// TIA Portal project "环氧乙烷灭菌器（XG2-C）260909_V18" (V18)

(* hardware
DEVICE "S7-1200 station_1"  S7-1200 Station
   slot 0: "Rack_0"  S7-1200 Rack  Rack  V1.0
   slot 1: "PLC_1"  CPU 1214C DC/DC/DC  6ES7 214-1AG40-0XB0  V4.2
   slot 2: "DI 8x24VDC_1"  6ES7 221-1BF32-0XB0  V2.0
   slot 3: "DQ 8x24VDC _1"  SM 1222 DQ8 x 24VDC  6ES7 222-1BF32-0XB0  V2.0
   slot 4: "DQ 8x24VDC _2"  SM 1222 DQ8 x 24VDC  6ES7 222-1BF32-0XB0  V2.0
   slot 5: "AI 4xRTD_1"  SM 1231 AI4 x RTD  6ES7 231-5PD32-0XB0  V2.0
   slot 6: "AI 4x13BIT_1"  6ES7 231-4HD32-0XB0  V2.0
*)

// ===== PLC "PLC_1"  CPU 1214C DC/DC/DC =====
// protected blocks, not shown: "0程序运行控制流程", "1预处理", "2保压", "3加湿", "4加药", "5灭菌", "6脉动", "7通风", "Main", "紧急脉动", "紧急通风"

VAR_GLOBAL   // PLC tag table "默认变量表"
   "Clock_Byte" AT %MB0 : Byte;
   "Clock_10Hz" AT %M0.0 : Bool;
   "Clock_5Hz" AT %M0.1 : Bool;
   "Clock_2.5Hz" AT %M0.2 : Bool;
   "Clock_2Hz" AT %M0.3 : Bool;
   "Clock_1.25Hz" AT %M0.4 : Bool;
   "Clock_1Hz" AT %M0.5 : Bool;
   "Clock_0.625Hz" AT %M0.6 : Bool;
   "Clock_0.5Hz" AT %M0.7 : Bool;
   "System_Byte" AT %MB1 : Byte;
   "FirstScan" AT %M1.0 : Bool;
   "DiagStatusUpdate" AT %M1.1 : Bool;
   "AlwaysTRUE" AT %M1.2 : Bool;
   "AlwaysFALSE" AT %M1.3 : Bool;
   "回空阀" AT %Q0.0 : Bool;
   "空" AT %IW64 : Int;
   "空(1)" AT %IW66 : Int;
   "催化前温度" AT %IW112 : Int;
   "催化后温度" AT %IW114 : Int;
   "内室压力P1" AT %IW160 : Int;
   "内室压力P2" AT %IW162 : Int;
   "内室湿度" AT %IW164 : Int;
   "前加湿阀" AT %Q0.1 : Bool;
   "后加湿阀" AT %Q0.2 : Bool;
   "加药阀关" AT %Q0.5 : Bool;
   "开装载门" AT %Q0.6 : Bool;
   "关装载门" AT %Q0.7 : Bool;
   "加热系统断电-脱扣器" AT %Q1.0 : Bool;
   "空压机" AT %Q1.1 : Bool;
   "开卸载门" AT %Q3.0 : Bool;
   "关卸载门" AT %Q3.1 : Bool;
   "卸载门加热" AT %Q3.2 : Bool;
   "运行灯" AT %Q3.3 : Bool;
   "待机灯" AT %Q3.4 : Bool;
   "报警灯" AT %Q3.5 : Bool;
   "快抽空阀2" AT %Q3.6 : Bool;
   "真空泵2" AT %Q3.7 : Bool;
   "快抽空阀" AT %Q0.3 : Bool;
   "加药阀开" AT %Q0.4 : Bool;
   "前门脚踢开关" AT %I0.0 : Bool;
   "前门开位" AT %I0.1 : Bool;
   "前门关位" AT %I0.2 : Bool;
   "前门障碍" AT %I0.3 : Bool;
   "前门电机过载" AT %I0.4 : Bool;
   "穿刺气缸穿刺位" AT %I0.5 : Bool;
   "下水位" AT %I0.6 : Bool;
   "压缩气压力检测" AT %I0.7 : Bool;
   "急停按钮" AT %I1.0 : Bool;
   "空压机保护" AT %I1.1 : Bool;
   "真空泵保护" AT %I1.2 : Bool;
   "真空泵2保护" AT %I1.3 : Bool;
   "排气压力开关" AT %I1.4 : Bool;
   "水箱上水位" AT %I1.5 : Bool;
   "后门开位" AT %I2.0 : Bool;
   "后门关位" AT %I2.1 : Bool;
   "后门障碍" AT %I2.2 : Bool;
   "后门脚踢开关" AT %I2.3 : Bool;
   "后门电机过载" AT %I2.4 : Bool;
   "后门开门按钮" AT %I2.5 : Bool;
   "后门关门按钮" AT %I2.6 : Bool;
   "关机确认信号" AT %I2.7 : Bool;
   "真空泵1" AT %Q2.0 : Bool;
   "蜂鸣器" AT %Q2.1 : Bool;
   "前部加热" AT %Q2.2 : Bool;
   "后部加热" AT %Q2.3 : Bool;
   "装载门加热" AT %Q2.4 : Bool;
   "汽化器加热" AT %Q2.5 : Bool;
   "慢抽空阀" AT %Q2.6 : Bool;
   "加热供电" AT %Q2.7 : Bool;
   "运行灯-蓝色" AT %Q4.0 : Bool;
   "待机灯-白灯" AT %Q4.1 : Bool;
   "报警灯-红灯" AT %Q4.2 : Bool;
   "预留" AT %Q4.3 : Bool;
   "预留(1)" AT %Q4.4 : Bool;
   "预留(2)" AT %Q4.5 : Bool;
   "预留(3)" AT %Q4.6 : Bool;
   "预留(4)" AT %Q4.7 : Bool;
   "前部温度" AT %IW128 : Int;
   "后部温度" AT %IW130 : Int;
   "前门温度" AT %IW132 : Int;
   "内室温度1" AT %IW134 : Int;
   "仿真秒沿" AT %M100.0 : Bool;
   "Tag_2" AT %M2.0 : Bool;
   "运行程序时间清零" AT %M5.0 : Bool;
   "汽化器温度" AT %IW166 : Int;
   "Tag_3" AT %M100.1 : Bool;
   "Tag_4" AT %M1.7 : Bool;
   "Tag_5" AT %MW102 : Hw_Device;
END_VAR

DATA_BLOCK "双泵控制_DB"   // DB142
{ S7_Optimized_Access := 'TRUE' }
VERSION : 0.1
// stored: InstanceOfName 双泵控制
"双泵控制"
BEGIN
END_DATA_BLOCK

DATA_BLOCK "单扉组态"   // DB160
{ S7_Optimized_Access := 'TRUE' }
VERSION : 0.1
   VAR
      Configuration : Struct
         Block_length : USInt := 16;
         Block_ID : USInt := 196;
         "Version" : USInt := 5;
         Subversion : USInt;
         Slot_1 : USInt := 1;
         Slot_2 : USInt := 255;   // 原组态插槽2的模块 没有了
         Slot_3 : USInt := 2;   // 原组态插槽3的模块去了 插槽2按照顺序排
         Slot_4 : USInt := 255;   // 原组态插槽4的模块 没有了
         Slot_5 : USInt := 3;   // 原组态插槽5的模块 去了插槽3 按照顺序排
         Slot_6 : USInt := 4;   // 原组态插槽6的模块 去了插槽4 按照顺序排
         Slot_7 : USInt := 255;
         Slot_8 : USInt := 255;
         Slot_9 : USInt := 255;
         Slot_101 : USInt := 255;
         Slot_102 : USInt := 255;
         Slot_103 : USInt := 255;
      END_STRUCT;
   END_VAR
BEGIN
END_DATA_BLOCK

DATA_BLOCK "双扉组态"   // DB161
{ S7_Optimized_Access := 'TRUE' }
VERSION : 0.1
   VAR
      Configuration : Struct
         Block_length : USInt := 16;
         Block_ID : USInt := 196;
         "Version" : USInt := 5;
         Subversion : USInt;
         Slot_1 : USInt := 1;
         Slot_2 : USInt := 2;
         Slot_3 : USInt := 3;
         Slot_4 : USInt := 4;
         Slot_5 : USInt := 5;
         Slot_6 : USInt := 6;
         Slot_7 : USInt := 255;
         Slot_8 : USInt := 255;
         Slot_9 : USInt := 255;
         Slot_101 : USInt := 255;
         Slot_102 : USInt := 255;
         Slot_103 : USInt := 255;
      END_STRUCT;
   END_VAR
BEGIN
END_DATA_BLOCK

DATA_BLOCK "单扉双泵组态"   // DB162
{ S7_Optimized_Access := 'TRUE' }
VERSION : 0.1
   VAR
      Configuration : Struct
         Block_length : USInt := 16;
         Block_ID : USInt := 196;
         "Version" : USInt := 5;
         Subversion : USInt;
         Slot_1 : USInt := 1;
         Slot_2 : USInt := 255;   // 原组态插槽2的模块 没有了
         Slot_3 : USInt := 2;   // 原组态插槽3的模块去了 插槽2按照顺序排
         Slot_4 : USInt := 3;   // 原组态插槽4的模块 没有了
         Slot_5 : USInt := 4;   // 原组态插槽5的模块 去了插槽3 按照顺序排
         Slot_6 : USInt := 5;   // 原组态插槽6的模块 去了插槽4 按照顺序排
         Slot_7 : USInt := 255;
         Slot_8 : USInt := 255;
         Slot_9 : USInt := 255;
         Slot_101 : USInt := 255;
         Slot_102 : USInt := 255;
         Slot_103 : USInt := 255;
      END_STRUCT;
   END_VAR
BEGIN
END_DATA_BLOCK

// folder: 100数据参数汇总

DATA_BLOCK "触摸屏"   // DB48
{ S7_Optimized_Access := 'FALSE' }
VERSION : 0.1
   VAR
      设备配置 : Word;
      选择程序 : Word;
      程序类型 : Word;
      手动操作1 : Word;
      手动操作2 : Word;
      维护类报警A1 : Word;
      维护类报警A2 : Word;
      维护类报警A3 : Word;
      门机构报警B1 : Word;
      门机构报警B2 : Word;
      启动类报警C1 : Word;
      启动类报警C2 : Word;
      全局类报警E1 : Word;
      全局类报警E2 : Word;
      全局类报警E3 : Word;
      运行错误报警F1 : Word;
      运行错误报警F2 : Word;
      运行错误报警F3 : Word;
      REO报警内容R1 : Word;
      REO报警内容R2 : Word;
      追溯类报警 : Word;
      维护类报警A1开关 : Word;
      维护类报警A2开关 : Word;
      维护类报警A3开关 : Word;
      门机构报警B1开关 : Word;
      门机构报警B2开关 : Word;
      启动类报警C1开关 : Word;
      启动类报警C2开关 : Word;
      全局类报警E1开关 : Word;
      全局类报警E2开关 : Word;
      全局类报警E3开关 : Word;
      运行错误报警F1开关 : Word;
      运行错误报警F2开关 : Word;
      运行错误报警F3开关 : Word;
      内室压力上传HMI : Int;
      内室温度上传HMI : Int;
      内室湿度上传HMI : Int;
      标志位1 : Word;
      标志位2 : Word;
      预留8 : Word;
      按钮1 : Word;
      按钮2 : Word;
      按钮3 : Word;
      按钮4 : Word;
      DI空压机保护 : Bool;
      DI真空泵保护 : Bool;
      DI前门电机过载 : Bool;
      DI前门脚踢开关 : Bool;
      DI后门脚踢开关 : Bool;
      DI排气压力开关 : Bool;
      DI关机确认信号 : Bool;
      DI前门开位 : Bool;
      DI前门关位 : Bool;
      DI前门障碍 : Bool;
      DI穿刺气缸位 : Bool;
      DI水箱上水位 : Bool;
      DI水箱下水位 : Bool;
      DI压缩气压力检测 : Bool;
      DI真空泵2保护 : Bool;
      DI后门开位 : Bool;
      DI后门关位 : Bool;
      DI后门障碍 : Bool;
      DI急停按钮 : Bool;
      DI后门电机过载 : Bool;
      DI空压机过载信号 : Bool;
      DI真空泵1过载信号 : Bool;
      DI真空泵2过载信号 : Bool;
      DI开后门按钮 : Bool;
      DI关后门按钮 : Bool;
      DI预留1 : Bool;
      DI预留2 : Bool;
      DI预留3 : Bool;
      DI预留4 : Bool;
      DI预留5 : Bool;
      DI预留6 : Bool;
      DI预留7 : Bool;
      DO回空阀 : Bool;
      DO前加湿阀 : Bool;
      DO后加湿阀 : Bool;
      DO快抽空阀 : Bool;
      DO加药阀开 : Bool;
      DO加药阀关 : Bool;
      DO慢抽空阀 : Bool;
      DO_2 : Bool;
      DO_1 : Bool;
      DO加热供电 : Bool;
      DO运行灯 : Bool;
      DO待机灯 : Bool;
      DO报警灯 : Bool;
      DO蜂鸣器 : Bool;
      DO腔体加热系统断电 : Bool;
      DO开装载门 : Bool;
      DO关装载门 : Bool;
      DO开卸载门 : Bool;
      DO关卸载门 : Bool;
      DO前部加热 : Bool;
      DO后部加热 : Bool;
      DO装载门加热 : Bool;
      DO卸载门加热 : Bool;
      DO汽化器加热 : Bool;
      DO_5 : Bool;
      DO_4 : Bool;
      "DO" : Bool;
      DO_3 : Bool;
      DO真空泵1 : Bool;
      DO真空泵2 : Bool;
      DO关机确认 : Bool;
      DO快抽空阀2 : Bool;
      DO空压机 : Bool;
      DO预留1 : Bool;
      DO预留2 : Bool;
      DO预留3 : Bool;
      DO预留4 : Bool;
      DO预留5 : Bool;
      DO预留6 : Bool;
      DO预留7 : Bool;
      DO预留8 : Bool;
      DO预留9 : Bool;
      DO预留10 : Bool;
      DO预留11 : Bool;
      DO预留12 : Bool;
      DO预留13 : Bool;
      DO预留14 : Bool;
      DO预留15 : Bool;
      追溯报警缓存 : Word;
      预留15 : Word;
      预留16 : Word;
      预留17 : Word;
      预留18 : Word;
      预留19 : Word;
      预留20 : Word;
      L抽空限度 : Int;
      L预热时间 : Int;
      L保压时间 : Int;
      L泄露率 : Int;
      L加湿湿度 : Int;
      "L加湿压力上限（没用到该变量）" : Int;
      L加湿均匀时间 : Int;
      L灭菌压力回压下限 : Int;
      L灭菌压力上限 : Int;
      L灭菌时间 : Int;
      L脉动次数 : Int;
      L脉动上限 : Int;
      L脉动下限 : Int;
      L通风上限 : Int;
      L通风下限 : Int;
      L通风时间 : Int;
      L结束时间 : Int;
      L灭菌温度 : Int;
      L加药平衡时间 : Int;
      L加湿湿化最短时间 : Int;
      "L加湿湿化让步10%时间" : Int;
      "L加湿湿化让步15%时间" : Int;
      "L最低湿度让步时间（湿度＞40%）" : Int;
      L预处理抽空预估时间 : Int;
      L加湿回空预估时间 : Int;
      L加湿抽空预估时间 : Int;
      L加药上升预估时间 : Int;
      L单次脉动时间 : Int;
      L紧急脉动次数 : Int;
      L紧急通风时间 : Int;
      备用 : Int;
      备用_1 : Int;
      备用_2 : Int;
      备用_3 : Int;
      L腔体前部控制温度 : Int;
      L腔体后部控制温度 : Int;
      L前门控制温度 : Int;
      "L后部控制温度（参数无用）" : Int;
      L加湿汽化控制温度 : Int;
      L加药汽化控制温度 : Int;
      L前部控温上偏差 : Int;
      L前部控温下偏差 : Int;
      L后部控温上偏差 : Int;
      L后部控温下偏差 : Int;
      L前门控温上偏差 : Int;
      L前门控温下偏差 : Int;
      L加湿汽化控温上偏差 : Int;
      L加湿汽化控温下偏差 : Int;
      L加药汽化控温上偏差 : Int;
      L加药汽化控温下偏差 : Int;
      L抽空超时报警时间 : Int;
      L回空超时报警时间 : Int;
      L加湿超时报警时间 : Int;
      L灭菌压力低报警时间 : Int;
      L腔体前部升温超时 : Int;
      L腔体后部升温超时 : Int;
      L门升温超时 : Int;
      L汽化器升温超时 : Int;
      L前部超温温度 : Int;
      L后部超温温度 : Int;
      L门超温温度 : Int;
      L加湿汽化超温温度 : Int;
      L加药汽化超温温度 : Int;
      L加药时间上限 : Int;
      L后门控制温度 : Int;
      L后门控温上限 : Int;
      L后门控温下限 : Int;
      L催化箱控制温度 : Int;
      L催化箱控制温度上限 : Int;
      L催化箱升温超时报警时间 : Int;
      L机壳报警温度 : Int;
      L通风阶段解毒时间 : Int;
      L脉动提前加热时间 : Int;
      L催化前超温报警温度 : Int;
      L催化后超温报警温度 : Int;
      L灭菌后回空至大气压偏差值 : Int;
      L慢排阀抽空下限 : Int;
      备用_4 : Int;
      备用_5 : Int;
      备用_6 : Int;
      H抽空限度 : Int;
      H预热时间 : Int;
      H保压时间 : Int;
      H泄露率 : Int;
      H加湿湿度 : Int;
      "H加湿压力上限(没用到该变量)" : Int;
      H加湿均匀时间 : Int;
      H灭菌压力回压下限 : Int;
      H灭菌压力上限 : Int;
      H灭菌时间 : Int;
      H脉动次数 : Int;
      H脉动上限 : Int;
      H脉动下限 : Int;
      H通风上限 : Int;
      H通风下限 : Int;
      H通风时间 : Int;
      H结束时间 : Int;
      H灭菌温度 : Int;
      H加药平衡时间 : Int;
      H加湿湿化最短时间 : Int;
      "H加湿湿化让步10%时间" : Int;
      "H加湿湿化让步15%时间" : Int;
      "H最低湿度让步时间(湿度＞40%)" : Int;
      H预处理抽空预估时间 : Int;
      H加湿回空预估时间 : Int;
      H加湿抽空预估时间 : Int;
      H加药上升预估时间 : Int;
      H单次脉动时间 : Int;
      H紧急脉动次数 : Int;
      H紧急通风时间 : Int;
      备用_7 : Int;
      备用_8 : Int;
      备用_9 : Int;
      备用_10 : Int;
      H腔体前部控制温度 : Int;
      H腔体后部控制温度 : Int;
      H前门控制温度 : Int;
      "H后部控制温度(参数无用)" : Int;
      H加湿汽化控制温度 : Int;
      H加药汽化控制温度 : Int;
      H前部控温上偏差 : Int;
      H前部控温下偏差 : Int;
      H后部控温上偏差 : Int;
      H后部控温下偏差 : Int;
      H前门控温上偏差 : Int;
      H前门控温下偏差 : Int;
      H加湿汽化控温上偏差 : Int;
      H加湿汽化控温下偏差 : Int;
      H加药汽化控温上偏差 : Int;
      H加药汽化控温下偏差 : Int;
      H抽空超时报警时间 : Int;
      H回空超时报警时间 : Int;
      H加湿超时报警时间 : Int;
      H灭菌压力低报警时间 : Int;
      H腔体前部升温超时 : Int;
      H腔体后部升温超时 : Int;
      H门升温超时 : Int;
      H汽化器升温超时 : Int;
      H前部超温温度 : Int;
      H后部超温温度 : Int;
      H门超温温度 : Int;
      H加湿汽化超温温度 : Int;
      H加药汽化超温温度 : Int;
      H加药时间上限 : Int;
      H后门控制温度 : Int;
      H后门控温上限 : Int;
      H后门控温下限 : Int;
      H催化箱控制温度 : Int;
      H催化箱控制温度上限 : Int;
      H催化箱升温超时报警时间 : Int;
      H机壳报警温度 : Int;
      H通风阶段解毒时间 : Int;
      H脉动提前加热时间 : Int;
      H催化前超温报警温度 : Int;
      H催化后超温报警温度 : Int;
      H灭菌后回空至大气压偏差值 : Int;
      H慢排阀抽空下限 : Int;
      备用_11 : Int;
      备用_12 : Int;
      备用_13 : Int;
      保压运行结果 : Int;
      程序编辑选择 : Int;
      门状态 : Int;
      程序运行编号 : Int;
      程序运行大阶段 : Int;
      程序运行小阶段 : Int;
      手动退出提示 : Int;
      运行结果 : Int;
      "总时间运行值-小时" : Int;
      "总时间运行值-分钟" : Int;
      "总时间运行值-秒钟" : Int;
      "大阶段时间运行值-小时" : Int;
      "大阶段时间运行值-分钟" : Int;
      "大阶段时间运行值-秒钟" : Int;
      "运行时间倒计时-小时" : Int;
      "运行时间倒计时-分钟" : Int;
      "运行时间倒计时-秒" : Int;
      运行百分比 : Int;
      Static_8 : Int;
      小阶段运行时间分 : Int;
      小阶段运行时间秒 : Int;
      Static_7 : Int;
      Static_11 : Int;
      脉动运行次数 : Int;
      "预处理运行时间（min）" : Int;
      "保压运行时间（min）" : Int;
      "加湿运行时间（min）" : Int;
      "加药运行时间（min）" : Int;
      "灭菌运行时间（min）" : Int;
      "脉动运行时间（min）" : Int;
      "通风阶段运行时间（min）" : Int;
      "结束运行时间（min）" : Int;
      "紧急脉动时间（min）" : Int;
      "紧急通风时间（min）" : Int;
      Static_3 : Int;
      预处理最高温度 : Int;
      预处理最低温度 : Int;
      预处理最高压力 : Int;
      预处理最低压力 : Int;
      预处理最高湿度 : Int;
      预处理最低湿度 : Int;
      保压最高温度 : Int;
      保压最低温度 : Int;
      保压最高压力 : Int;
      保压最低压力 : Int;
      保压最高湿度 : Int;
      保压最低湿度 : Int;
      加湿最高温度 : Int;
      加湿最低温度 : Int;
      加湿最高压力 : Int;
      加湿最低压力 : Int;
      加湿最高湿度 : Int;
      加湿最低湿度 : Int;
      加药最高温度 : Int;
      加药最低温度 : Int;
      加药最高压力 : Int;
      加药最低压力 : Int;
      加药最高湿度 : Int;
      加药最低湿度 : Int;
      灭菌最高温度 : Int;
      灭菌最低温度 : Int;
      灭菌最高压力 : Int;
      灭菌最低压力 : Int;
      灭菌最高湿度 : Int;
      灭菌最低湿度 : Int;
      脉动最高温度 : Int;
      脉动最低温度 : Int;
      脉动最高压力 : Int;
      脉动最低压力 : Int;
      脉动最高湿度 : Int;
      脉动最低湿度 : Int;
      通风最高温度 : Int;
      通风最低温度 : Int;
      通风最高压力 : Int;
      通风最低压力 : Int;
      通风最高湿度 : Int;
      通风最低湿度 : Int;
      紧急脉动最高压力 : Int;
      紧急脉动最低压力 : Int;
      紧急通风最高压力 : Int;
      紧急通风最低压力 : Int;
      水位状态 : Int;
      气罐状态 : Int;
      预热名称显示 : Int;
      预处理阶段预估值 : Int;
      保压阶段预估值 : Int;
      加湿阶段预估值 : Int;
      进药阶段预估值 : Int;
      灭菌阶段预估值 : Int;
      脉动阶段预估值 : Int;
      通风阶段预估值 : Int;
      结束阶段预估值 : Int;
      紧急脉动预估时间 : Int;
      紧急通风预估时间 : Int;
      异常退出回空预估时间 : Int;
      程序总计时时 : Int;
      程序总计时分 : Int;
      程序总计时秒 : Int;
      大阶段计时时 : Int;
      大阶段计时分 : Int;
      大阶段计时秒 : Int;
      小阶段计时时 : Int;
      小阶段计时分 : Int;
      小阶段计时秒 : Int;
      "预处理运行时间（秒）" : Int;
      "保压运行时间（秒）" : Int;
      "加湿运行时间（秒）" : Int;
      "加药运行时间（秒）" : Int;
      "灭菌运行时间（秒）" : Int;
      "脉动运行时间（秒）" : Int;
      "通风阶段运行时间（秒）" : Int;
      "结束运行时间（秒）" : Int;
      "紧急脉动时间（秒）" : Int;
      "紧急通风时间（秒）" : Int;
      前门加热膜最大加热时间秒 : Int;
      汽化器最大加热时间秒 : Int;
      后门加热膜最大加热时间秒 : Int;
      "压缩气最大恢复时间 秒" : Int;
      "加药最长时间（从穿刺到压力稳定）秒" : Int;
      "加湿完成最长时间 分钟" : Int;
      "抽空最大时间 秒" : Int;
      "回空最大时间 秒" : Int;
      新屏内1环百分比 : Int;
      新屏内2环百分比 : Int;
      新屏内3环百分比 : Int;
      新屏最外环百分比 : Int;
      打印数据标志 : Int;
      预留_1 : Int;
      预留_2 : Int;
      预留_3 : Int;
      预留_4 : Int;
      预留_5 : Int;
      预留_6 : Int;
      预留_7 : Int;
      预留_8 : Int;
      内室温度1偏差校准 : Int;
      内室温度2偏差校准 : Int;
      前部温度偏差校准 : Int;
      后部温度偏差校准 : Int;
      前门温度偏差校准 : Int;
      汽化温度偏差校准 : Int;
      Static_6 : Int;
      内室湿度偏差校准 : Int;
      内室压力1偏差校准 : Int;
      内室压力2偏差校准 : Int;
      Static_1 : Int;
      Static_2 : Int;
      催化前温度偏差校准 : Int;
      催化后温度偏差校准 : Int;
      后门温度偏差校准 : Int;
      备用偏差校准 : Int;
      备用偏差校准_1 : Int;
      "年  设置" : Int;
      "月  设置" : Int;
      "日  设置" : Int;
      "时  设置" : Int;
      "分  设置" : Int;
      "秒  设置" : Int;
      "星期几  设置" : Int;
      "年     显示" : Int;
      "月  显示" : Int;
      "日  显示" : Int;
      "时  显示" : Int;
      "分  显示" : Int;
      "秒  显示" : Int;
      网络模式 : Int;
      内室温度1 : Int;
      内室温度2 : Int;
      前部温度 : Int;
      后部温度 : Int;
      前门温度 : Int;
      汽化温度 : Int;
      无 : Int;
      内室湿度 : Int;
      内室压力P1 : Int;
      内室压力P2 : Int;
      稀释管路压力 : Int;
      催化箱保护温度 : Int;
      催化前温度 : Int;
      催化后温度 : Int;
      后门温度 : Int;
      界面地址 : Int;
      设备型号 : Int;
      设备容积 : Int;
      打印模式选择 : Int;
      PLC程序版本1 : Int;
      PLC程序版本2 : Int;
      PLC程序版本3 : Int;
      PLC程序版本4 : Int;
      PLC程序版本5 : Int;
      PLC程序版本6 : Int;
      PLC程序版本7 : Int;
      PLC程序版本8 : Int;
      本地大气压 : Int;
      开门压差 : Int;
      回空压差 : Int;
      Static_4 : Int;
      Static_5 : Int;
      催化剂寿命 : Int;
      结束后自动开门最大时间间隔 : Int;
      程序结束自动脉动时间 : Int;
      前部升温超时报警时间 : Int;
      后部升温超时报警时间 : Int;
      前门升温超时报警时间 : Int;
      汽化器升温超时报警时间 : Int;
      后门升温超时报警时间 : Int;
      启动内室温度下偏差 : Int;
      启动非内室温度下偏差 : Int;
      慢排阀开启间隔 : Int;
      慢排阀关闭间隔 : Int;
      慢排阀间歇控制脉动次数 : Int;
      解毒器慢排阀开启脉动次数 : Int;
      程序结束后自动开门 : Int;
      催化箱升温超时报警时间 : Int;
      门动作时间上限 : Int;
      预留_9 : Int;
      预留_10 : Int;
      数据存储间隔 : Int;
      催化剂使用时间 : Int;
      本地大气压设置值 : Int;
      IP一段 : Int;
      IP二段 : Int;
      IP三段 : Int;
      IP四段 : Int;
      网关一段 : Int;
      网关二段 : Int;
      网关三段 : Int;
      网关四段 : Int;
      子网掩码一段 : Int;
      子网掩码二段 : Int;
      子网掩码三段 : Int;
      子网掩码四段 : Int;
      "上次保养日期(年)" : Int;
      "上次保养日期(月)" : Int;
      "上次保养日期(日)" : Int;
      "下次保养日期(年)" : Int;
      "下次保养日期(月)" : Int;
      "下次保养日期(日)" : Int;
      计划保养周期天数 : Int := 180;
      上次保养次数 : Int;
      距离上次保养天数 : Int;
      距离上次保养循环次数 : Int;
      计划保养循环次数 : Int := 180;
      总运行次数 : Int;
      已完成次数 : Int;
      未完成次数 : Int;
      结束蜂鸣器开启时间 : Int;
      结束蜂鸣器关闭时间 : Int;
      结束蜂鸣器鸣响时间 : Int;
      报警蜂鸣器开启时间 : Int;
      报警蜂鸣器关闭时间 : Int;
      报警蜂鸣器鸣响时间 : Int;
      预留_12 : Int;
      预留_13 : Int;
      预留_14 : Int;
      预留_15 : Int;
      设备编号12 : Int;
      设备编号34 : Int;
      设备编号56 : Int;
      设备编号78 : Int;
      用户地址 : Int;
      权限地址 : Int;
      紧急脉动打印标志 : Int;
      泄漏率 : Int;
      语言切换 : Int;
      正使用泵的编号 : Int;
      预处理打印间隔 : Int;
      保压打印间隔 : Int;
      加湿打印间隔 : Int;
      加药打印间隔 : Int;
      灭菌打印间隔 : Int;
      脉动打印间隔 : Int;
      通风打印间隔 : Int;
      灭菌曲线打印间隔 : Int;
      通风曲线打印间隔 : Int;
      "其他阶段 曲线打印间隔" : Int;
      触摸屏用曲线打印间隔设定值 : Int;
      预留_37 : Int;
      预留_38 : Int;
      预留_39 : Int;
      预留_40 : Int;
      预留_41 : Int;
      预留_42 : Int;
      预留_43 : Int;
      预留_44 : Int;
   END_VAR
BEGIN
END_DATA_BLOCK

DATA_BLOCK "默认参数"   // DB1000
{ S7_Optimized_Access := 'FALSE' }
VERSION : 0.1
   VAR
      L抽空限度 : Int := 180;
      L预热时间 : Int := 20;
      L保压时间 : Int := 20;
      L泄露率 : Int := 1;
      L加湿湿度 : Int := 600;
      "L加湿压力上限（没用到该变量）" : Int := 220;
      L加湿均匀时间 : Int := 20;
      L灭菌压力回压下限 : Int := 350;
      L灭菌压力上限 : Int := 800;
      L灭菌时间 : Int := 180;
      L脉动次数 : Int := 5;
      L脉动上限 : Int := 750;
      L脉动下限 : Int := 180;
      L通风上限 : Int := 750;
      L通风下限 : Int := 300;
      L通风时间 : Int := 1320;
      L结束时间 : Int := 2;
      L灭菌温度 : Int := 370;
      L加药平衡时间 : Int := 5;
      L加湿湿化最短时间 : Int := 30;
      "L加湿湿化让步10%时间" : Int := 40;
      "L加湿湿化让步15%时间" : Int := 50;
      "L最低湿度让步时间（湿度＞40%）" : Int := 60;
      L预处理抽空预估时间 : Int := 4;
      L加湿回空预估时间 : Int := 1;
      L加湿抽空预估时间 : Int := 4;
      L加药上升预估时间 : Int := 2;
      L单次脉动时间 : Int := 6;
      L紧急脉动次数 : Int := 5;
      L紧急通风时间 : Int := 150;
      L本地大气压设定 : Int := 1010;
      备用_1 : Int;
      备用_2 : Int;
      备用_3 : Int;
      L腔体前部控制温度 : Int := 375;
      L腔体后部控制温度 : Int := 375;
      L前门控制温度 : Int := 375;
      "L后部控制温度（参数无用）" : Int := 375;
      L加湿汽化控制温度 : Int := 1100;
      L加药汽化控制温度 : Int := 700;
      L前部控温上偏差 : Int := 5;
      L前部控温下偏差 : Int := -5;
      L后部控温上偏差 : Int := 5;
      L后部控温下偏差 : Int := -5;
      L前门控温上偏差 : Int := 5;
      L前门控温下偏差 : Int := -5;
      L加湿汽化控温上偏差 : Int := 50;
      L加湿汽化控温下偏差 : Int := -10;
      L加药汽化控温上偏差 : Int := 20;
      L加药汽化控温下偏差 : Int := 0;
      L抽空超时报警时间 : Int := 15;
      L回空超时报警时间 : Int := 8;
      L加湿超时报警时间 : Int := 90;
      L灭菌压力低报警时间 : Int := 5;
      L腔体前部升温超时 : Int := 90;
      L腔体后部升温超时 : Int := 90;
      L门升温超时 : Int := 90;
      L汽化器升温超时 : Int := 10;
      L前部超温温度 : Int := 50;
      L后部超温温度 : Int := 50;
      L门超温温度 : Int := 50;
      L加湿汽化超温温度 : Int := 200;
      L加药汽化超温温度 : Int := 200;
      L加药时间上限 : Int := 10;
      L后门控制温度 : Int := 375;
      L后门控温上限 : Int := 5;
      L后门控温下限 : Int := -5;
      L催化箱控制温度 : Int := 2650;
      L催化箱控制温度上限 : Int := 50;
      L催化箱升温超时报警时间 : Int := 60;
      L机壳报警温度 : Int := 600;
      L通风阶段解毒时间 : Int := 120;
      L脉动提前加热时间 : Int := 60;
      L催化前超温报警温度 : Int := 3800;
      L催化后超温报警温度 : Int := 4200;
      L灭菌后回空至大气压偏差值 : Int;
      L慢排阀抽空下限 : Int;
      备用_4 : Int;
      备用_5 : Int;
      备用_6 : Int;
      H抽空限度 : Int := 180;
      H预热时间 : Int := 20;
      H保压时间 : Int := 20;
      H泄露率 : Int := 1;
      H加湿湿度 : Int := 600;
      "H加湿压力上限(没用到该变量)" : Int := 220;
      H加湿均匀时间 : Int := 20;
      H灭菌压力回压下限 : Int := 350;
      H灭菌压力上限 : Int := 800;
      H灭菌时间 : Int := 60;
      H脉动次数 : Int := 5;
      H脉动上限 : Int := 750;
      H脉动下限 : Int := 180;
      H通风上限 : Int := 750;
      H通风下限 : Int := 300;
      H通风时间 : Int := 720;
      H结束时间 : Int := 2;
      H灭菌温度 : Int := 550;
      H加药平衡时间 : Int := 5;
      H加湿湿化最短时间 : Int := 30;
      "H加湿湿化让步10%时间" : Int := 40;
      "H加湿湿化让步15%时间" : Int := 50;
      "H最低湿度让步时间(湿度＞40%)" : Int := 60;
      H预处理抽空预估时间 : Int := 4;
      H加湿回空预估时间 : Int := 1;
      H加湿抽空预估时间 : Int := 4;
      H加药上升预估时间 : Int := 2;
      H单次脉动时间 : Int := 6;
      H紧急脉动次数 : Int := 5;
      H紧急通风时间 : Int := 150;
      H本地大气压设定 : Int := 1010;
      备用_8 : Int := 0;
      备用_9 : Int := 0;
      备用_10 : Int := 0;
      H腔体前部控制温度 : Int := 560;
      H腔体后部控制温度 : Int := 560;
      H前门控制温度 : Int := 560;
      "H后部控制温度(参数无用)" : Int := 560;
      H加湿汽化控制温度 : Int := 1100;
      H加药汽化控制温度 : Int := 700;
      H前部控温上偏差 : Int := 5;
      H前部控温下偏差 : Int := -5;
      H后部控温上偏差 : Int := 5;
      H后部控温下偏差 : Int := -5;
      H前门控温上偏差 : Int := 5;
      H前门控温下偏差 : Int := -5;
      H加湿汽化控温上偏差 : Int := 50;
      H加湿汽化控温下偏差 : Int := -10;
      H加药汽化控温上偏差 : Int := 20;
      H加药汽化控温下偏差 : Int := 0;
      H抽空超时报警时间 : Int := 15;
      H回空超时报警时间 : Int := 8;
      H加湿超时报警时间 : Int := 90;
      H灭菌压力低报警时间 : Int := 5;
      H腔体前部升温超时 : Int := 90;
      H腔体后部升温超时 : Int := 90;
      H门升温超时 : Int := 90;
      H汽化器升温超时 : Int := 10;
      H前部超温温度 : Int := 50;
      H后部超温温度 : Int := 50;
      H门超温温度 : Int := 50;
      H加湿汽化超温温度 : Int := 200;
      H加药汽化超温温度 : Int := 200;
      H加药时间上限 : Int := 10;
      H后门控制温度 : Int := 560;
      H后门控温上限 : Int := 5;
      H后门控温下限 : Int := -5;
      H催化箱控制温度 : Int := 2650;
      H催化箱控制温度上限 : Int := 50;
      H催化箱升温超时报警时间 : Int := 60;
      H机壳报警温度 : Int := 600;
      H通风阶段解毒时间 : Int := 120;
      H脉动提前加热时间 : Int := 60;
      H催化前超温报警温度 : Int := 3800;
      H催化后超温报警温度 : Int := 4200;
      H灭菌后回空至大气压偏差值 : Int := 0;
      H慢排阀抽空下限 : Int := 0;
      备用_11 : Int := 0;
      备用_12 : Int := 0;
      备用_13 : Int := 0;
      备用_14 : Int;
      备用_15 : Int;
      备用_16 : Int;
      备用_17 : Int;
      备用_18 : Int;
      备用_19 : Int;
      备用_20 : Int;
      本地大气压 : Int := 1010;
      开门压差 : Int := 50;
      回空压差 : Int := 20;
      Static_1 : Int := 0;
      Static_2 : Int := 0;
      催化剂寿命 : Int := 8000;
      结束后自动开门最大时间间隔 : Int := 600;
      程序结束自动脉动时间 : Int := 900;
      前部升温超时报警时间 : Int := 60;
      后部升温超时报警时间 : Int := 60;
      前门升温超时报警时间 : Int := 100;
      汽化器升温超时报警时间 : Int := 40;
      后门升温超时报警时间 : Int := 60;
      启动内室温度下偏差 : Int := 50;
      启动非内室温度下偏差 : Int := 100;
      慢排阀开启间隔 : Int := 0;
      慢排阀关闭间隔 : Int := 0;
      慢排阀间歇控制脉动次数 : Int := 0;
      解毒器慢排阀开启脉动次数 : Int := 3;
      程序结束后自动开门 : Int := 0;
      催化箱升温超时报警时间 : Int := 60;
      门动作时间上限 : Int := 39;
      预留_9 : Int;
      预留_10 : Int;
      预留_11 : Int;
      预留 : Int;
      预留_1 : Int;
      预留_2 : Int;
      预留_3 : Int;
      预留_4 : Int;
      YG抽空限度 : Int := 180;
      YG预热时间 : Int := 0;
      YG保压时间 : Int := 20;
      YG泄露率 : Int := 1;
      YG加湿湿度 : Int := 0;
      "YG加湿压力上限（没用到该变量）" : Int := 220;
      YG加湿均匀时间 : Int := 0;
      YG灭菌压力回压下限 : Int := 350;
      YG灭菌压力上限 : Int := 800;
      YG灭菌时间 : Int := 0;
      YG脉动次数 : Int := 5;
      YG脉动上限 : Int := 750;
      YG脉动下限 : Int := 180;
      YG通风上限 : Int := 750;
      YG通风下限 : Int := 300;
      YG通风时间 : Int := 150;
      YG结束时间 : Int := 2;
      YG灭菌温度 : Int := 370;
      YG加药平衡时间 : Int := 0;
      YG加湿湿化最短时间 : Int := 0;
      "YG加湿湿化让步10%时间" : Int := 10;
      "YG加湿湿化让步15%时间" : Int := 20;
      "YG最低湿度让步时间（湿度＞40%）" : Int := 30;
      YG预处理抽空预估时间 : Int := 4;
      YG加湿回空预估时间 : Int := 1;
      YG加湿抽空预估时间 : Int := 4;
      YG加药上升预估时间 : Int := 2;
      YG单次脉动时间 : Int := 6;
      YG紧急脉动次数 : Int := 5;
      YG紧急通风时间 : Int := 150;
      YG本地大气压设定 : Int := 1010;
      备用_7 : Int := 0;
      备用_21 : Int := 0;
      备用_22 : Int := 0;
      YG腔体前部控制温度 : Int := 375;
      YG腔体后部控制温度 : Int := 375;
      YG前门控制温度 : Int := 375;
      "YG后部控制温度（参数无用）" : Int := 375;
      YG加湿汽化控制温度 : Int := 1100;
      YG加药汽化控制温度 : Int := 700;
      YG前部控温上偏差 : Int := 5;
      YG前部控温下偏差 : Int := -5;
      YG后部控温上偏差 : Int := 5;
      YG后部控温下偏差 : Int := -5;
      YG前门控温上偏差 : Int := 5;
      YG前门控温下偏差 : Int := -5;
      YG加湿汽化控温上偏差 : Int := 50;
      YG加湿汽化控温下偏差 : Int := -10;
      YG加药汽化控温上偏差 : Int := 20;
      YG加药汽化控温下偏差 : Int := 0;
      YG抽空超时报警时间 : Int := 15;
      YG回空超时报警时间 : Int := 8;
      YG加湿超时报警时间 : Int := 90;
      YG灭菌压力低报警时间 : Int := 5;
      YG腔体前部升温超时 : Int := 90;
      YG腔体后部升温超时 : Int := 90;
      YG门升温超时 : Int := 90;
      YG汽化器升温超时 : Int := 10;
      YG前部超温温度 : Int := 50;
      YG后部超温温度 : Int := 50;
      YG门超温温度 : Int := 50;
      YG加湿汽化超温温度 : Int := 200;
      YG加药汽化超温温度 : Int := 200;
      YG加药时间上限 : Int := 10;
      YG后门控制温度 : Int := 375;
      YG后门控温上限 : Int := 5;
      YG后门控温下限 : Int := -5;
      YG催化箱控制温度 : Int := 2650;
      YG催化箱控制温度上限 : Int := 50;
      YG催化箱升温超时报警时间 : Int := 60;
      YG机壳报警温度 : Int := 600;
      YG通风阶段解毒时间 : Int := 120;
      YG脉动提前加热时间 : Int := 60;
      YG催化前超温报警温度 : Int := 3800;
      YG催化后超温报警温度 : Int := 4200;
      YG灭菌后回空至大气压偏差值 : Int := 0;
      YG慢排阀抽空下限 : Int := 0;
      备用_23 : Int := 0;
      备用_24 : Int := 0;
      备用_25 : Int := 0;
      XL抽空限度 : Int := 180;
      XL预热时间 : Int := 0;
      XL保压时间 : Int := 20;
      XL泄露率 : Int := 1;
      XL加湿湿度 : Int := 600;
      "XL加湿压力上限（没用到该变量）" : Int := 220;
      XL加湿均匀时间 : Int := 0;
      XL灭菌压力回压下限 : Int := 350;
      XL灭菌压力上限 : Int := 800;
      XL灭菌时间 : Int := 0;
      XL脉动次数 : Int := 5;
      XL脉动上限 : Int := 750;
      XL脉动下限 : Int := 180;
      XL通风上限 : Int := 750;
      XL通风下限 : Int := 300;
      XL通风时间 : Int := 0;
      XL结束时间 : Int := 2;
      XL灭菌温度 : Int := 370;
      XL加药平衡时间 : Int := 5;
      XL加湿湿化最短时间 : Int := 30;
      "XL加湿湿化让步10%时间" : Int := 40;
      "XL加湿湿化让步15%时间" : Int := 50;
      "XL最低湿度让步时间（湿度＞40%）" : Int := 60;
      XL预处理抽空预估时间 : Int := 4;
      XL加湿回空预估时间 : Int := 1;
      XL加湿抽空预估时间 : Int := 4;
      XL加药上升预估时间 : Int := 2;
      XL单次脉动时间 : Int := 6;
      XL紧急脉动次数 : Int := 5;
      XL紧急通风时间 : Int := 150;
      XL本地大气压设定 : Int := 1010;
      备用_26 : Int := 0;
      备用_27 : Int := 0;
      备用_28 : Int := 0;
      XL腔体前部控制温度 : Int := 375;
      XL腔体后部控制温度 : Int := 375;
      XL前门控制温度 : Int := 375;
      "XL后部控制温度（参数无用）" : Int := 375;
      XL加湿汽化控制温度 : Int := 1100;
      XL加药汽化控制温度 : Int := 700;
      XL前部控温上偏差 : Int := 5;
      XL前部控温下偏差 : Int := -5;
      XL后部控温上偏差 : Int := 5;
      XL后部控温下偏差 : Int := -5;
      XL前门控温上偏差 : Int := 5;
      XL前门控温下偏差 : Int := -5;
      XL加湿汽化控温上偏差 : Int := 50;
      XL加湿汽化控温下偏差 : Int := -10;
      XL加药汽化控温上偏差 : Int := 20;
      XL加药汽化控温下偏差 : Int := 0;
      XL抽空超时报警时间 : Int := 15;
      XL回空超时报警时间 : Int := 8;
      XL加湿超时报警时间 : Int := 90;
      XL灭菌压力低报警时间 : Int := 5;
      XL腔体前部升温超时 : Int := 90;
      XL腔体后部升温超时 : Int := 90;
      XL门升温超时 : Int := 90;
      XL汽化器升温超时 : Int := 10;
      XL前部超温温度 : Int := 50;
      XL后部超温温度 : Int := 50;
      XL门超温温度 : Int := 50;
      XL加湿汽化超温温度 : Int := 200;
      XL加药汽化超温温度 : Int := 200;
      XL加药时间上限 : Int := 10;
      XL后门控制温度 : Int := 375;
      XL后门控温上限 : Int := 5;
      XL后门控温下限 : Int := -5;
      XL催化箱控制温度 : Int := 2650;
      XL催化箱控制温度上限 : Int := 50;
      XL催化箱升温超时报警时间 : Int := 60;
      XL机壳报警温度 : Int := 600;
      XL通风阶段解毒时间 : Int := 120;
      XL脉动提前加热时间 : Int := 60;
      XL催化前超温报警温度 : Int := 3800;
      XL催化后超温报警温度 : Int := 4200;
      XL灭菌后回空至大气压偏差值 : Int := 0;
      XL慢排阀抽空下限 : Int := 0;
      备用_29 : Int := 0;
      备用_30 : Int := 0;
      备用_31 : Int := 0;
   END_VAR
BEGIN
END_DATA_BLOCK

// folder: 101中间变量

DATA_BLOCK "中间变量"   // DB3
{ S7_Optimized_Access := 'FALSE' }
VERSION : 0.1
   VAR
      启动内室温度下限 : Int;
      启动内室温度上限 : Int;
      启动前部温度下限 : Int;
      启动后部温度下限 : Int;
      启动门温度下限 : Int;
      启动前部温度上限 : Int;
      启动后部温度上限 : Int;
      启动门温度上限 : Int;
      脉动次数 : Int;
      加药DJS时间 : Int;
      测试设定值2 : Int;
      腔体前部超温报警上限 : Int;
      腔体后部超温报警上限 : Int;
      前门超温报警上限 : Int;
      汽化器超温报警上限 : Int;
      内室温度超温报警上限 : Int;
      两压力差值 : Int;
      腔体前部持续加热时间 : Int;
      腔体后部持续加热时间 : Int;
      前门持续加热时间 : Int;
      汽化器持续加热时间 : Int;
      后门持续加热时间 : Int;
      催化箱持续加热时间 : Int;
      预处理大阶段运行时间分 : Int;
      预处理大阶段运行时间秒 : Int;
      预处理小阶段运行时间分 : Int;
      预处理小阶段运行时间秒 : Int;
      预处理小阶段名称 : Int;
      预处理真空泵1输出 : Bool;
      预处理快抽空阀V4输出 : Bool;
      Static_2 : Bool;
      Static_3 : Bool;
      预处理加药阀关输出 : Bool;
      加湿加药阀关输出 : Bool;
      保压大阶段运行时间分 : Int;
      保压大阶段运行时间秒 : Int;
      保压小阶段运行时间分 : Int;
      保压小阶段运行时间秒 : Int;
      保压小阶段名称 : Int;
      Static_4 : Bool;
      保压加药阀关输出 : Bool;
      Static_7 : Bool;
      加湿大阶段运行时间分 : Int;
      加湿大阶段运行时间秒 : Int;
      加湿小阶段运行时间分 : Int;
      加湿小阶段运行时间秒 : Int;
      加湿小阶段名称 : Int;
      Static_5 : Bool;
      加湿真空泵1输出 : Bool;
      加湿快抽空阀V4输出 : Bool;
      加湿回空阀输出 : Bool;
      前加湿阀V2输出 : Bool;
      后加湿阀V3输出 : Bool;
      加药阶段V5阀开输出 : Bool;
      加药阶段V11阀输出 : Bool;
      加药大阶段运行时间分 : Int;
      加药大阶段运行时间秒 : Int;
      加药小阶段运行时间分 : Int;
      加药小阶段运行时间秒 : Int;
      加药小阶段名称 : Int;
      灭菌大阶段运行时间分 : Int;
      灭菌大阶段运行时间秒 : Int;
      灭菌小阶段运行时间分 : Int;
      灭菌小阶段运行时间秒 : Int;
      灭菌小阶段名称 : Int;
      脉动大阶段运行时间分 : Int;
      脉动大阶段运行时间秒 : Int;
      脉动小阶段运行时间分 : Int;
      脉动小阶段运行时间秒 : Int;
      脉动小阶段名称 : Int;
      脉动阶段回空阀V1输出 : Bool;
      脉动阶段快抽空阀V4输出 : Bool;
      脉动阶段慢抽空阀V8输出 : Bool;
      脉动阶段真空泵1输出 : Bool;
      脉动阶段解毒稀释V9输出 : Bool;
      脉动阶段解毒阀V10输出 : Bool;
      通风真空泵1输出 : Bool;
      通风大阶段运行时间分 : Int;
      通风大阶段运行时间秒 : Int;
      通风小阶段运行时间分 : Int;
      通风小阶段运行时间秒 : Int;
      通风小阶段名称 : Int;
      通风阶段回空阀V1输出 : Bool;
      通风阶段快抽空阀V4输出 : Bool;
      结束阶段回空阀V1输出 : Bool;
      程序正常结束标志 : Bool;
      加药阶段V5阀关输出 : Bool;
      灭菌阶段V5阀关输出 : Bool;
      脉动阶段V5阀关输出 : Bool;
      通风阶段V5阀关输出 : Bool;
      结束大阶段运行时间分 : Int;
      结束大阶段运行时间秒 : Int;
      结束小阶段运行时间分 : Int;
      结束小阶段运行时间秒 : Int;
      结束小阶段名称 : Int;
      紧急脉动大阶段运行时间分 : Int;
      紧急脉动大阶段运行时间秒 : Int;
      紧急脉动小阶段运行时间分 : Int;
      紧急脉动小阶段运行时间秒 : Int;
      紧急脉动小阶段名称 : Int;
      紧急通风大阶段运行时间分 : Int;
      紧急通风大阶段运行时间秒 : Int;
      紧急通风小阶段运行时间分 : Int;
      紧急通风小阶段运行时间秒 : Int;
      紧急通风小阶段名称 : Int;
      预留_10 : Int;
      DJS预处理 : Int;
      DJS保压 : Int;
      DJS加湿 : Int;
      DJS加药 : Int;
      DJS灭菌 : Int;
      DJS脉动 : Int;
      DJS通风 : Int;
      DJS结束 : Int;
      DJS紧急脉动 : Int;
      DJS紧急通风 : Int;
      开门脉动小阶段 : Int;
      已经进行过脉动标志 : Int;
      程序结束15分钟标志位 : Int;
      催化加热1标志 : Bool;
      催化加热2标志 : Bool;
      催化箱加热标志 : Bool;
      汽化器加热标志 : Bool;
      前部加热标志 : Bool;
      后部加热标志 : Bool;
      前门加热标志 : Bool;
      后门加热标志 : Bool;
      内室工作压力 : Int;
      催化类报警开V11标志 : Bool;
      程序报警退出标志 : Bool;
      紧急脉动真空泵1输出 : Bool;
      紧急脉动回空阀 : Bool;
      紧急脉动快抽阀 : Bool;
      紧急脉动直排阀 : Bool;
      Static_1 : Bool;
      程序暂停标志 : Bool;
      程序紧急通风标志 : Bool;
      紧急通风快抽空阀 : Bool;
      紧急通风回空阀 : Bool;
      紧急通风直排阀 : Bool;
      后门停止加热条件 : Bool;
      催化加热控制阶段热回收阀打开 : Bool;
      内室工作温度 : Int;
      维护类报警A1缓存 : Word;
      维护类报警A2缓存 : Word;
      维护类报警A3缓存 : Word;
      门机构报警B1缓存 : Word;
      门机构报警B2缓存 : Word;
      启动类报警C1缓存 : Word;
      启动类报警C2缓存 : Word;
      全局类报警E1缓存 : Word;
      全局类报警E2缓存 : Word;
      全局类报警E3缓存 : Word;
      运行错误报警F1缓存 : Word;
      运行错误报警F2缓存 : Word;
      运行错误报警F3缓存 : Word;
      蜂鸣器输出标志 : Bool;
      上电时间统计沿 : Bool;
      上电1秒标志 : Bool;
      上电5秒标志 : Bool;
      上电30秒标志 : Bool;
      上电60秒标志 : Bool;
      与REO通讯故障标志 : Bool;
      开门脉动快抽空阀V4 : Bool;
      开门脉动回空阀V1 : Bool;
      开门脉动真空泵 : Bool;
      结束灯自动 : Bool;
      沿预留_9 : Bool;
      沿预留_10 : Bool;
      沿预留_11 : Bool;
      沿预留_12 : Bool;
      沿预留_13 : Bool;
      上电时间统计 : Int;
      后门停止加热上限1 : Int;
      前门状态输出 : Int;
      后门状态输出 : Int;
      E014报警计算1 : Int;
      E014报警计算2 : Int;
      E014报警计算3 : Int;
      E014报警计算4 : Int;
      启动程序时有报警标志 : Bool;
      预热完成标志 : Bool;
      保压完成标志 : Bool;
      加湿完成标志 : Bool;
      加药完成标志 : Bool;
      灭菌完成标志 : Bool;
      脉动完成标志 : Bool;
      通风完成标志 : Bool;
      泄露测试完成标志 : Bool;
      紧急脉动完成标志 : Bool;
      紧急通风完成标志 : Bool;
      结束阶段完成标志 : Bool;
      预热阶段抽空超时报警 : Bool;
      保压阶段保压超时报警 : Bool;
      加湿阶段抽空超时报警 : Bool;
      加湿阶段加湿超时报警 : Bool;
      加药阶段加药失败报警 : Bool;
      加药阶段进药压力过高报警 : Bool;
      灭菌阶段压力过高报警 : Bool;
      脉动阶段抽空超时报警 : Bool;
      脉动阶段回空超时报警 : Bool;
      紧急通风真空泵1输出 : Bool;
      紧急情况阶段完成标志 : Bool;
      回空超时报警时间 : DInt;
      阶段最大压力 : Int;
      阶段最小压力 : Int;
      阶段最大湿度 : Int;
      阶段最小湿度 : Int;
      阶段最大温度 : Int;
      阶段最小温度 : Int;
      紧急脉动打印标志 : Int;
      加药平衡时间 : DInt;
      REO报警1缓存 : Word;
      REO报警2缓存 : Word;
      打印标志1 : Int;
      灭菌时间小于60分钟允许灭菌标志 : Bool;
      内室压力正常标志 : Bool;
      内室湿度正常标志 : Bool;
      内室温度正常标志 : Bool;
      双泵设备泵切换标志 : Bool;
      时钟冻结标志 : Bool;
      仿真标志 : Bool;
      预留bool3 : Bool;
      预留bool4 : Bool;
      预留bool5 : Bool;
      预留bool6 : Bool;
      预留bool7 : Bool;
      预留bool8 : Bool;
      预留bool9 : Bool;
      预留bool10 : Bool;
      预留bool11 : Bool;
      预处理最高温度 : Int;
      预处理最低温度 : Int;
      预处理最高压力 : Int;
      预处理最低压力 : Int;
      预处理最高湿度 : Int;
      预处理最低湿度 : Int;
      保压最高温度 : Int;
      保压最低温度 : Int;
      保压最高压力 : Int;
      保压最低压力 : Int;
      保压最高湿度 : Int;
      保压最低湿度 : Int;
      加湿最高温度 : Int;
      加湿最低温度 : Int;
      加湿最高压力 : Int;
      加湿最低压力 : Int;
      加湿最高湿度 : Int;
      加湿最低湿度 : Int;
      加药最高温度 : Int;
      加药最低温度 : Int;
      加药最高压力 : Int;
      加药最低压力 : Int;
      加药最高湿度 : Int;
      加药最低湿度 : Int;
      灭菌最高温度 : Int;
      灭菌最低温度 : Int;
      灭菌最高压力 : Int;
      灭菌最低压力 : Int;
      灭菌最高湿度 : Int;
      灭菌最低湿度 : Int;
      脉动最高温度 : Int;
      脉动最低温度 : Int;
      脉动最高压力 : Int;
      脉动最低压力 : Int;
      脉动最高湿度 : Int;
      脉动最低湿度 : Int;
      通风最高温度 : Int;
      通风最低温度 : Int;
      通风最高压力 : Int;
      通风最低压力 : Int;
      通风最高湿度 : Int;
      通风最低湿度 : Int;
      紧急脉动最高压力 : Int;
      紧急脉动最低压力 : Int;
      紧急通风最高压力 : Int;
      紧急通风最低压力 : Int;
      小阶段名称缓存 : Int;
      Dint值 : DInt;
      Int值 : Int;
   END_VAR
BEGIN
END_DATA_BLOCK

DATA_BLOCK "中间转换变量_DB"   // DB70
{ S7_Optimized_Access := 'TRUE' }
VERSION : 0.1
// stored: InstanceOfName 中间转换变量
"中间转换变量"
BEGIN
END_DATA_BLOCK

// folder: 12门功能控制

DATA_BLOCK "前门控制逻辑_DB"   // DB27
{ S7_Optimized_Access := 'TRUE' }
VERSION : 0.1
// stored: InstanceOfName 门控制逻辑
"门控制逻辑"
BEGIN
END_DATA_BLOCK

DATA_BLOCK "后门控制逻辑_DB"   // DB28
{ S7_Optimized_Access := 'TRUE' }
VERSION : 0.1
// stored: InstanceOfName 门控制逻辑
"门控制逻辑"
BEGIN
END_DATA_BLOCK

DATA_BLOCK "门功能控制_DB"   // DB102
{ S7_Optimized_Access := 'TRUE' }
VERSION : 0.1
// stored: InstanceOfName 门功能控制
"门功能控制"
BEGIN
END_DATA_BLOCK

DATA_BLOCK "程序结束自动开门_DB"   // DB136
{ S7_Optimized_Access := 'TRUE' }
VERSION : 0.1
// stored: InstanceOfName 程序结束自动开门
"程序结束自动开门"
BEGIN
END_DATA_BLOCK

DATA_BLOCK "程序结束长时间不开门自动脉动_DB"   // DB145
{ S7_Optimized_Access := 'TRUE' }
VERSION : 0.1
// stored: InstanceOfName 程序结束长时间不开门自动脉动
"程序结束长时间不开门自动脉动"
BEGIN
END_DATA_BLOCK

// folder: 14加热功能控制

DATA_BLOCK "加热功能控制_DB"   // DB103
{ S7_Optimized_Access := 'TRUE' }
VERSION : 0.1
// stored: InstanceOfName 加热功能控制
"加热功能控制"
BEGIN
END_DATA_BLOCK

// folder: 17页面控制

DATA_BLOCK "页面跳转控制_DB"   // DB104
{ S7_Optimized_Access := 'TRUE' }
VERSION : 0.1
// stored: InstanceOfName 页面跳转控制
"页面跳转控制"
BEGIN
END_DATA_BLOCK

// folder: 200尾气处理器

DATA_BLOCK "尾气处理器"   // DB1
{ S7_Optimized_Access := 'FALSE' }
VERSION : 0.1
   VAR
      处理器输入映像区 : Word;
      处理器输出映像区 : Word;
      处理器风速传感器 : Int;
      处理器房间浓度传感器 : Int;
      处理器催化后浓度传感器 : Int;
      处理器催化前温度 : Int;
      处理器催化后温度 : Int;
      处理器机壳温度 : Int;
      处理器报警内容1 : Word;
      处理器报警内容2 : Word;
      处理器大阶段 : Int;
      "处理器大阶段运行时间-时" : Int;
      "处理器大阶段运行时间-分" : Int;
      "处理器大阶段运行时间-秒" : Int;
      处理器风机运行总时间 : DInt;
      处理器催化剂已使用时间 : Int;
      处理器运行次数 : Int;
      处理器软件版本号01 : Word;
      处理器软件版本号23 : Word;
      处理器软件版本号45 : Word;
      处理器软件版本号67 : Word;
      处理器软件版本号89 : Word;
      处理器软件版本号1011 : Word;
      处理器软件版本号1213 : Word;
      处理器软件版本号1415 : Word;
      处理器心跳信号 : Int;
      处理器信息预留1 : Word;
      处理器信息预留2 : Word;
      处理器信息预留3 : Word;
      处理器信息预留4 : Word;
      处理器信息预留5 : Word;
      处理器信息预留6 : Word;
      处理器信息预留7 : Word;
      处理器信息预留8 : Word;
      处理器信息预留9 : Word;
      处理器信息预留10 : Word;
      处理器信息预留11 : Word;
      处理器信息预留12 : Word;
      处理器信息预留13 : Word;
      处理器信息预留14 : Word;
      处理器信息预留15 : Word;
      处理器信息预留16 : Word;
      处理器信息预留17 : Word;
      处理器信息预留18 : Word;
      处理器信息预留19 : Word;
      处理器信息预留20 : Word;
      处理器信息预留21 : Word;
      处理器信息预留22 : Word;
      处理器信息预留23 : Word;
      灭菌器1手动操作 : Word;
      灭菌器1报警开关1 : Word;
      灭菌器1报警开关2 : Word;
      灭菌器1按钮 : Word;
      灭菌器1大阶段 : Int;
      灭菌器1要处理器进行的阶段 : Int;
      灭菌器1信息预留0 : Int;
      灭菌器1信息预留1 : Int;
      灭菌器1信息预留2 : Int;
      灭菌器1信息预留3 : Int;
      灭菌器1催化前控制温度 : Int;
      灭菌器1催化前控温上限偏差 : Int;
      灭菌器1催化前控温下限偏差 : Int;
      灭菌器1催化前超温报警温度 : Int;
      灭菌器1催化后超温报警温度 : Int;
      灭菌器1待机温度 : Int;
      灭菌器1待机上偏差 : Int;
      灭菌器1待机下偏差 : Int;
      灭菌器1升温超时报警时间 : Int;
      灭菌器1冷却时间 : Int;
      灭菌器1机壳报警温度 : Int;
      灭菌器1冷却超时报警时间 : Int;
      灭菌器1风机运行最低报警风速 : Int;
      灭菌器1催化剂设定寿命 : Int;
      灭菌器1催化前温度偏差校准 : Int;
      灭菌器1催化后温度偏差校准 : Int;
      灭菌器1机壳温度偏差校准 : Int;
      灭菌器1风速传感器偏差校准 : Int;
      灭菌器1房间浓度传感器偏差校准 : Int;
      灭菌器1催化后浓度传感器偏差校准 : Int;
      灭菌器1报警蜂鸣器频率开时间 : Int;
      灭菌器1报警蜂鸣器频率关时间 : Int;
      灭菌器1报警蜂鸣器蜂鸣时间 : Int;
      灭菌器1心跳信号 : Int;
      灭菌器1灭菌提前加热时间 : Int;
      灭菌器1通风催化处理时间 : Int;
      灭菌器1信息预留6 : Int;
      灭菌器1信息预留7 : Int;
      灭菌器1信息预留8 : Int;
      灭菌器1信息预留9 : Int;
      灭菌器1信息预留10 : Int;
      灭菌器1信息预留11 : Int;
      灭菌器1信息预留12 : Int;
      灭菌器1信息预留13 : Int;
      灭菌器1信息预留14 : Int;
      灭菌器1信息预留15 : Int;
      灭菌器1信息预留16 : Int;
      灭菌器1信息预留17 : Int;
      灭菌器1信息预留18 : Int;
      灭菌器1信息预留19 : Int;
      灭菌器2大阶段 : Int;
      灭菌器2要处理器进行的阶段 : Int;
      灭菌器2心跳信号 : Int;
      灭菌器2信息预留0 : Int;
      灭菌器2信息预留1 : Int;
      灭菌器2信息预留2 : Int;
      灭菌器2信息预留3 : Int;
      灭菌器2信息预留4 : Int;
      灭菌器2信息预留5 : Int;
      灭菌器2信息预留6 : Int;
      灭菌器2信息预留7 : Int;
      灭菌器2信息预留8 : Int;
      灭菌器2信息预留9 : Int;
      灭菌器2信息预留10 : Int;
      灭菌器2信息预留11 : Int;
   END_VAR
BEGIN
END_DATA_BLOCK

DATA_BLOCK "尾气处理器处理_DB"   // DB91
{ S7_Optimized_Access := 'TRUE' }
VERSION : 0.1
// stored: InstanceOfName 尾气处理器处理
"尾气处理器处理"
BEGIN
END_DATA_BLOCK

// folder: 21蜂鸣器控制

DATA_BLOCK "蜂鸣器控制流程子程序_DB"   // DB97
{ S7_Optimized_Access := 'TRUE' }
VERSION : 0.1
// stored: InstanceOfName 蜂鸣器控制流程子程序
"蜂鸣器控制流程子程序"
BEGIN
END_DATA_BLOCK

// folder: 3报警处理

DATA_BLOCK "报警处理_DB"   // DB99
{ S7_Optimized_Access := 'TRUE' }
VERSION : 0.1
// stored: InstanceOfName 报警处理
"报警处理"
BEGIN
END_DATA_BLOCK

// folder: 4网络设置

DATA_BLOCK "网络设置IP路由地址"   // DB143
{ S7_Optimized_Access := 'FALSE' }
VERSION : 0.1
   VAR
      IP_config : Struct
         Header : IF_CONF_Header;
         IPdata : IF_CONF_v4;
      END_STRUCT;
   END_VAR
BEGIN
   IP_config.Header.SubfieldCount := 1;
   IP_config.IPdata.Mode := 1;
   IP_config.IPdata.InterfaceAddress.ADDR[1] := 192;
   IP_config.IPdata.InterfaceAddress.ADDR[2] := 168;
   IP_config.IPdata.InterfaceAddress.ADDR[3] := 0;
   IP_config.IPdata.InterfaceAddress.ADDR[4] := 2;
   IP_config.IPdata.SubnetMask.ADDR[1] := 255;
   IP_config.IPdata.SubnetMask.ADDR[2] := 255;
   IP_config.IPdata.SubnetMask.ADDR[3] := 255;
   IP_config.IPdata.SubnetMask.ADDR[4] := 0;
   IP_config.IPdata.DefaultRouter.ADDR[1] := 192;
   IP_config.IPdata.DefaultRouter.ADDR[2] := 168;
   IP_config.IPdata.DefaultRouter.ADDR[3] := 0;
   IP_config.IPdata.DefaultRouter.ADDR[4] := 1;
END_DATA_BLOCK

DATA_BLOCK "网络设置IP路由地址默认"   // DB150
{ S7_Optimized_Access := 'TRUE' }
VERSION : 0.1
   VAR
      IP_config : Struct
         Header : IF_CONF_Header;
         IPdata : IF_CONF_v4;
      END_STRUCT;
   END_VAR
BEGIN
   IP_config.Header.SubfieldCount := 1;
   IP_config.IPdata.Mode := 1;
   IP_config.IPdata.InterfaceAddress.ADDR[1] := 192;
   IP_config.IPdata.InterfaceAddress.ADDR[2] := 168;
   IP_config.IPdata.InterfaceAddress.ADDR[3] := 0;
   IP_config.IPdata.InterfaceAddress.ADDR[4] := 2;
   IP_config.IPdata.SubnetMask.ADDR[1] := 255;
   IP_config.IPdata.SubnetMask.ADDR[2] := 255;
   IP_config.IPdata.SubnetMask.ADDR[3] := 255;
   IP_config.IPdata.SubnetMask.ADDR[4] := 0;
   IP_config.IPdata.DefaultRouter.ADDR[1] := 192;
   IP_config.IPdata.DefaultRouter.ADDR[2] := 168;
   IP_config.IPdata.DefaultRouter.ADDR[3] := 0;
   IP_config.IPdata.DefaultRouter.ADDR[4] := 1;
END_DATA_BLOCK

DATA_BLOCK "新网络设置_DB"   // DB151
{ S7_Optimized_Access := 'TRUE' }
VERSION : 0.1
// stored: InstanceOfName 新网络设置
"新网络设置"
BEGIN
END_DATA_BLOCK

// folder: 5智慧屏功能

DATA_BLOCK "智慧屏功能_DB"   // DB89
{ S7_Optimized_Access := 'TRUE' }
VERSION : 0.1
// stored: InstanceOfName 智慧屏功能
"智慧屏功能"
BEGIN
END_DATA_BLOCK

// folder: 6系统设置

DATA_BLOCK "系统参数设置_DB"   // DB100
{ S7_Optimized_Access := 'TRUE' }
VERSION : 0.1
// stored: InstanceOfName 系统参数设置
"系统参数设置"
BEGIN
END_DATA_BLOCK

// folder: 7程序参数

DATA_BLOCK "参数转换变量"   // DB2
{ S7_Optimized_Access := 'FALSE' }
VERSION : 0.1
   VAR
      M抽空限度 : Int;
      M预热时间 : Int;
      M保压时间 : Int;
      M泄露率 : Int;
      M加湿湿度 : Int;
      "M加湿压力上限（没用到该变量）" : Int;
      M加湿均匀时间 : Int;
      M灭菌压力回压下限 : Int;
      M灭菌压力上限 : Int;
      M灭菌时间 : Int;
      M脉动次数 : Int;
      M脉动上限 : Int;
      M脉动下限 : Int;
      M通风上限 : Int;
      M通风下限 : Int;
      M通风时间 : Int;
      M结束时间 : Int;
      M灭菌温度 : Int;
      M加药平衡时间 : Int;
      M加湿湿化最短时间 : Int;
      "M加湿湿化让步10%时间" : Int;
      "M加湿湿化让步15%时间" : Int;
      "M最低湿度让步时间（湿度＞40%）" : Int;
      M预处理抽空预估时间 : Int;
      M加湿回空预估时间 : Int;
      M加湿抽空预估时间 : Int;
      M加药上升预估时间 : Int;
      M单次脉动时间 : Int;
      M紧急脉动次数 : Int;
      M紧急通风时间 : Int;
      M本地大气压设定 : Int;
      备用_1 : Int;
      备用_2 : Int;
      备用_3 : Int;
      M腔体前部控制温度 : Int;
      M腔体后部控制温度 : Int;
      M前门控制温度 : Int;
      "M后部控制温度（参数无用）" : Int;
      M加湿汽化控制温度 : Int;
      M加药汽化控制温度 : Int;
      M前部控温上偏差 : Int;
      M前部控温下偏差 : Int;
      M后部控温上偏差 : Int;
      M后部控温下偏差 : Int;
      M前门控温上偏差 : Int;
      M前门控温下偏差 : Int;
      M加湿汽化控温上偏差 : Int;
      M加湿汽化控温下偏差 : Int;
      M加药汽化控温上偏差 : Int;
      M加药汽化控温下偏差 : Int;
      M抽空超时报警时间 : Int;
      M回空超时报警时间 : Int;
      M加湿超时报警时间 : Int;
      M灭菌压力低报警时间 : Int;
      M腔体前部升温超时 : Int;
      M腔体后部升温超时 : Int;
      M门升温超时 : Int;
      M汽化器升温超时 : Int;
      M前部超温温度 : Int;
      M后部超温温度 : Int;
      M门超温温度 : Int;
      M加湿汽化超温温度 : Int;
      M加药汽化超温温度 : Int;
      M加药时间上限 : Int;
      M后门控制温度 : Int;
      M后门控温上限 : Int;
      M后门控温下限 : Int;
      M催化箱控制温度 : Int;
      M催化箱控制温度上限 : Int;
      M催化箱升温超时报警时间 : Int;
      M机壳报警温度 : Int;
      M通风阶段解毒时间 : Int;
      M脉动提前加热时间 : Int;
      M催化前超温报警温度 : Int;
      M催化后超温报警温度 : Int;
      M灭菌后回空至大气压偏差值 : Int;
      M慢排阀抽空下限 : Int;
      备用_4 : Int;
      备用_5 : Int;
      备用_6 : Int;
   END_VAR
BEGIN
END_DATA_BLOCK

DATA_BLOCK "参数恢复默认_DB"   // DB10
{ S7_Optimized_Access := 'TRUE' }
VERSION : 0.1
// stored: InstanceOfName 参数恢复默认
"参数恢复默认"
BEGIN
END_DATA_BLOCK

DATA_BLOCK "程序运行参数传递_DB"   // DB85
{ S7_Optimized_Access := 'TRUE' }
VERSION : 0.1
// stored: InstanceOfName 程序运行参数传递
"程序运行参数传递"
BEGIN
END_DATA_BLOCK

DATA_BLOCK "2、药罐处理"   // DB109
{ S7_Optimized_Access := 'FALSE' }
VERSION : 0.1
   VAR
      YG抽空限度 : Int;
      YG预热时间 : Int;
      YG保压时间 : Int;
      YG泄露率 : Int;
      YG加湿湿度 : Int;
      "YG加湿压力上限（没用到该变量）" : Int;
      YG加湿均匀时间 : Int;
      YG灭菌压力回压下限 : Int;
      YG灭菌压力上限 : Int;
      YG灭菌时间 : Int;
      YG脉动次数 : Int;
      YG脉动上限 : Int;
      YG脉动下限 : Int;
      YG通风上限 : Int;
      YG通风下限 : Int;
      YG通风时间 : Int;
      YG结束时间 : Int;
      YG灭菌温度 : Int;
      YG加药平衡时间 : Int;
      YG加湿湿化最短时间 : Int;
      "YG加湿湿化让步10%时间" : Int;
      "YG加湿湿化让步15%时间" : Int;
      "YG最低湿度让步时间（湿度＞40%）" : Int;
      YG预处理抽空预估时间 : Int;
      YG加湿回空预估时间 : Int;
      YG加湿抽空预估时间 : Int;
      YG加药上升预估时间 : Int;
      YG单次脉动时间 : Int;
      YG紧急脉动次数 : Int;
      YG紧急通风时间 : Int;
      YG本地大气压设定 : Int;
      备用_7 : Int;
      备用_21 : Int;
      备用_22 : Int;
      YG腔体前部控制温度 : Int;
      YG腔体后部控制温度 : Int;
      YG前门控制温度 : Int;
      "YG后部控制温度（参数无用）" : Int;
      YG加湿汽化控制温度 : Int;
      YG加药汽化控制温度 : Int;
      YG前部控温上偏差 : Int;
      YG前部控温下偏差 : Int;
      YG后部控温上偏差 : Int;
      YG后部控温下偏差 : Int;
      YG前门控温上偏差 : Int;
      YG前门控温下偏差 : Int;
      YG加湿汽化控温上偏差 : Int;
      YG加湿汽化控温下偏差 : Int;
      YG加药汽化控温上偏差 : Int;
      YG加药汽化控温下偏差 : Int;
      YG抽空超时报警时间 : Int;
      YG回空超时报警时间 : Int;
      YG加湿超时报警时间 : Int;
      YG灭菌压力低报警时间 : Int;
      YG腔体前部升温超时 : Int;
      YG腔体后部升温超时 : Int;
      YG门升温超时 : Int;
      YG汽化器升温超时 : Int;
      YG前部超温温度 : Int;
      YG后部超温温度 : Int;
      YG门超温温度 : Int;
      YG加湿汽化超温温度 : Int;
      YG加药汽化超温温度 : Int;
      YG加药时间上限 : Int;
      YG后门控制温度 : Int;
      YG后门控温上限 : Int;
      YG后门控温下限 : Int;
      YG催化箱控制温度 : Int;
      YG催化箱控制温度上限 : Int;
      YG催化箱升温超时报警时间 : Int;
      YG机壳报警温度 : Int;
      YG通风阶段解毒时间 : Int;
      YG脉动提前加热时间 : Int;
      YG催化前超温报警温度 : Int;
      YG催化后超温报警温度 : Int;
      YG灭菌后回空至大气压偏差值 : Int;
      YG慢排阀抽空下限 : Int;
      备用_23 : Int;
      备用_24 : Int;
      备用_25 : Int;
   END_VAR
BEGIN
END_DATA_BLOCK

DATA_BLOCK "3、泄露测试"   // DB110
{ S7_Optimized_Access := 'FALSE' }
VERSION : 0.1
   VAR
      XL抽空限度 : Int;
      XL预热时间 : Int;
      XL保压时间 : Int;
      XL泄露率 : Int;
      XL加湿湿度 : Int;
      "XL加湿压力上限（没用到该变量）" : Int;
      XL加湿均匀时间 : Int;
      XL灭菌压力回压下限 : Int;
      XL灭菌压力上限 : Int;
      XL灭菌时间 : Int;
      XL脉动次数 : Int;
      XL脉动上限 : Int;
      XL脉动下限 : Int;
      XL通风上限 : Int;
      XL通风下限 : Int;
      XL通风时间 : Int;
      XL结束时间 : Int;
      XL灭菌温度 : Int;
      XL加药平衡时间 : Int;
      XL加湿湿化最短时间 : Int;
      "XL加湿湿化让步10%时间" : Int;
      "XL加湿湿化让步15%时间" : Int;
      "XL最低湿度让步时间（湿度＞40%）" : Int;
      XL预处理抽空预估时间 : Int;
      XL加湿回空预估时间 : Int;
      XL加湿抽空预估时间 : Int;
      XL加药上升预估时间 : Int;
      XL单次脉动时间 : Int;
      XL紧急脉动次数 : Int;
      XL紧急通风时间 : Int;
      XL本地大气压设定 : Int;
      备用_26 : Int;
      备用_27 : Int;
      备用_28 : Int;
      XL腔体前部控制温度 : Int;
      XL腔体后部控制温度 : Int;
      XL前门控制温度 : Int;
      "XL后部控制温度（参数无用）" : Int;
      XL加湿汽化控制温度 : Int;
      XL加药汽化控制温度 : Int;
      XL前部控温上偏差 : Int;
      XL前部控温下偏差 : Int;
      XL后部控温上偏差 : Int;
      XL后部控温下偏差 : Int;
      XL前门控温上偏差 : Int;
      XL前门控温下偏差 : Int;
      XL加湿汽化控温上偏差 : Int;
      XL加湿汽化控温下偏差 : Int;
      XL加药汽化控温上偏差 : Int;
      XL加药汽化控温下偏差 : Int;
      XL抽空超时报警时间 : Int;
      XL回空超时报警时间 : Int;
      XL加湿超时报警时间 : Int;
      XL灭菌压力低报警时间 : Int;
      XL腔体前部升温超时 : Int;
      XL腔体后部升温超时 : Int;
      XL门升温超时 : Int;
      XL汽化器升温超时 : Int;
      XL前部超温温度 : Int;
      XL后部超温温度 : Int;
      XL门超温温度 : Int;
      XL加湿汽化超温温度 : Int;
      XL加药汽化超温温度 : Int;
      XL加药时间上限 : Int;
      XL后门控制温度 : Int;
      XL后门控温上限 : Int;
      XL后门控温下限 : Int;
      XL催化箱控制温度 : Int;
      XL催化箱控制温度上限 : Int;
      XL催化箱升温超时报警时间 : Int;
      XL机壳报警温度 : Int;
      XL通风阶段解毒时间 : Int;
      XL脉动提前加热时间 : Int;
      XL催化前超温报警温度 : Int;
      XL催化后超温报警温度 : Int;
      XL灭菌后回空至大气压偏差值 : Int;
      XL慢排阀抽空下限 : Int;
      备用_29 : Int;
      备用_30 : Int;
      备用_31 : Int;
   END_VAR
BEGIN
END_DATA_BLOCK

DATA_BLOCK "1、37℃程序"   // DB111
{ S7_Optimized_Access := 'FALSE' }
VERSION : 0.1
   VAR
      L抽空限度 : Int;
      L预热时间 : Int;
      L保压时间 : Int;
      L泄露率 : Int;
      L加湿湿度 : Int;
      "L加湿压力上限（没用到该变量）" : Int;
      L加湿均匀时间 : Int;
      L灭菌压力回压下限 : Int;
      L灭菌压力上限 : Int;
      L灭菌时间 : Int;
      L脉动次数 : Int;
      L脉动上限 : Int;
      L脉动下限 : Int;
      L通风上限 : Int;
      L通风下限 : Int;
      L通风时间 : Int;
      L结束时间 : Int;
      L灭菌温度 : Int;
      L加药平衡时间 : Int;
      L加湿湿化最短时间 : Int;
      "L加湿湿化让步10%时间" : Int;
      "L加湿湿化让步15%时间" : Int;
      "L最低湿度让步时间（湿度＞40%）" : Int;
      L预处理抽空预估时间 : Int;
      L加湿回空预估时间 : Int;
      L加湿抽空预估时间 : Int;
      L加药上升预估时间 : Int;
      L单次脉动时间 : Int;
      L紧急脉动次数 : Int;
      L紧急通风时间 : Int;
      L本地大气压设定 : Int;
      备用_1 : Int;
      备用_2 : Int;
      备用_3 : Int;
      L腔体前部控制温度 : Int;
      L腔体后部控制温度 : Int;
      L前门控制温度 : Int;
      "L后部控制温度（参数无用）" : Int;
      L加湿汽化控制温度 : Int;
      L加药汽化控制温度 : Int;
      L前部控温上偏差 : Int;
      L前部控温下偏差 : Int;
      L后部控温上偏差 : Int;
      L后部控温下偏差 : Int;
      L前门控温上偏差 : Int;
      L前门控温下偏差 : Int;
      L加湿汽化控温上偏差 : Int;
      L加湿汽化控温下偏差 : Int;
      L加药汽化控温上偏差 : Int;
      L加药汽化控温下偏差 : Int;
      L抽空超时报警时间 : Int;
      L回空超时报警时间 : Int;
      L加湿超时报警时间 : Int;
      L灭菌压力低报警时间 : Int;
      L腔体前部升温超时 : Int;
      L腔体后部升温超时 : Int;
      L门升温超时 : Int;
      L汽化器升温超时 : Int;
      L前部超温温度 : Int;
      L后部超温温度 : Int;
      L门超温温度 : Int;
      L加湿汽化超温温度 : Int;
      L加药汽化超温温度 : Int;
      L加药时间上限 : Int;
      L后门控制温度 : Int;
      L后门控温上限 : Int;
      L后门控温下限 : Int;
      L催化箱控制温度 : Int;
      L催化箱控制温度上限 : Int;
      L催化箱升温超时报警时间 : Int;
      L机壳报警温度 : Int;
      L通风阶段解毒时间 : Int;
      L脉动提前加热时间 : Int;
      L催化前超温报警温度 : Int;
      L催化后超温报警温度 : Int;
      L灭菌后回空至大气压偏差值 : Int;
      L慢排阀抽空下限 : Int;
      备用_4 : Int;
      备用_5 : Int;
      备用_6 : Int;
   END_VAR
BEGIN
END_DATA_BLOCK

DATA_BLOCK "程序数据编辑、保存（55℃参数除外）_DB"   // DB112
{ S7_Optimized_Access := 'TRUE' }
VERSION : 0.1
// stored: InstanceOfName 程序数据编辑、保存（55℃参数除外）
"程序数据编辑、保存（55℃参数除外）"
BEGIN
END_DATA_BLOCK

// folder: 9程序运行控制流程

DATA_BLOCK "8结束_DB"   // DB77
{ S7_Optimized_Access := 'TRUE' }
VERSION : 0.1
// stored: InstanceOfName 8结束
"8结束"
BEGIN
END_DATA_BLOCK

// folder: System blocks/Program resources

DATA_BLOCK "保压大阶段时间统计"   // DB4
{ S7_Optimized_Access := 'TRUE' }
AUTHOR : Simatic
FAMILY : IEC
NAME : IEC_TMR
VERSION : 1.0
// stored: InstanceOfName IEC_TIMER
"IEC_TIMER"
BEGIN
END_DATA_BLOCK

DATA_BLOCK "灭菌阶段额外增加0.5秒"   // DB5
{ S7_Optimized_Access := 'TRUE' }
AUTHOR : Simatic
FAMILY : IEC
NAME : IEC_TMR
VERSION : 1.0
// stored: InstanceOfName IEC_TIMER
"IEC_TIMER"
BEGIN
END_DATA_BLOCK

DATA_BLOCK "压力超上限延时"   // DB6
{ S7_Optimized_Access := 'TRUE' }
AUTHOR : Simatic
FAMILY : IEC
NAME : IEC_TMR
VERSION : 1.0
// stored: InstanceOfName IEC_TIMER
"IEC_TIMER"
BEGIN
END_DATA_BLOCK

DATA_BLOCK "前加湿阀等待关断时间"   // DB7
{ S7_Optimized_Access := 'TRUE' }
AUTHOR : Simatic
FAMILY : IEC
NAME : IEC_TMR
VERSION : 1.0
// stored: InstanceOfName IEC_TIMER
"IEC_TIMER"
BEGIN
END_DATA_BLOCK

DATA_BLOCK "后加湿阀等待关断时间"   // DB8
{ S7_Optimized_Access := 'TRUE' }
AUTHOR : Simatic
FAMILY : IEC
NAME : IEC_TMR
VERSION : 1.0
// stored: InstanceOfName IEC_TIMER
"IEC_TIMER"
BEGIN
END_DATA_BLOCK

DATA_BLOCK "后加湿阀开启间隔计时"   // DB9
{ S7_Optimized_Access := 'TRUE' }
AUTHOR : Simatic
FAMILY : IEC
NAME : IEC_TMR
VERSION : 1.0
// stored: InstanceOfName IEC_TIMER
"IEC_TIMER"
BEGIN
END_DATA_BLOCK

DATA_BLOCK "穿刺维持计时"   // DB11
{ S7_Optimized_Access := 'TRUE' }
AUTHOR : Simatic
FAMILY : IEC
NAME : IEC_TMR
VERSION : 1.0
// stored: InstanceOfName IEC_TIMER
"IEC_TIMER"
BEGIN
END_DATA_BLOCK

DATA_BLOCK "穿刺回位等待计时"   // DB12
{ S7_Optimized_Access := 'TRUE' }
AUTHOR : Simatic
FAMILY : IEC
NAME : IEC_TMR
VERSION : 1.0
// stored: InstanceOfName IEC_TIMER
"IEC_TIMER"
BEGIN
END_DATA_BLOCK

DATA_BLOCK "加药平衡计时"   // DB13
{ S7_Optimized_Access := 'TRUE' }
AUTHOR : Simatic
FAMILY : IEC
NAME : IEC_TMR
VERSION : 1.0
// stored: InstanceOfName IEC_TIMER
"IEC_TIMER"
BEGIN
END_DATA_BLOCK

DATA_BLOCK "运行标志清零延时"   // DB14
{ S7_Optimized_Access := 'TRUE' }
AUTHOR : Simatic
FAMILY : IEC
NAME : IEC_TMR
VERSION : 1.0
// stored: InstanceOfName IEC_TIMER
"IEC_TIMER"
BEGIN
END_DATA_BLOCK

DATA_BLOCK "预处理大阶段时间统计"   // DB15
{ S7_Optimized_Access := 'TRUE' }
AUTHOR : Simatic
FAMILY : IEC
NAME : IEC_TMR
VERSION : 1.0
// stored: InstanceOfName IEC_TIMER
"IEC_TIMER"
BEGIN
END_DATA_BLOCK

DATA_BLOCK "异常结束标志延时1秒"   // DB17
{ S7_Optimized_Access := 'TRUE' }
AUTHOR : Simatic
FAMILY : IEC
NAME : IEC_TMR
VERSION : 1.0
// stored: InstanceOfName IEC_TIMER
"IEC_TIMER"
BEGIN
END_DATA_BLOCK

DATA_BLOCK "保压运行标志延时1秒"   // DB18
{ S7_Optimized_Access := 'TRUE' }
AUTHOR : Simatic
FAMILY : IEC
NAME : IEC_TMR
VERSION : 1.0
// stored: InstanceOfName IEC_TIMER
"IEC_TIMER"
BEGIN
END_DATA_BLOCK

DATA_BLOCK "37℃预热复位按钮"   // DB19
{ S7_Optimized_Access := 'TRUE' }
AUTHOR : Simatic
FAMILY : IEC
NAME : IEC_TMR
VERSION : 1.0
// stored: InstanceOfName IEC_TIMER
"IEC_TIMER"
BEGIN
END_DATA_BLOCK

DATA_BLOCK "保压正常结束大阶段延时"   // DB20
{ S7_Optimized_Access := 'TRUE' }
AUTHOR : Simatic
FAMILY : IEC
NAME : IEC_TMR
VERSION : 1.0
// stored: InstanceOfName IEC_TIMER
"IEC_TIMER"
BEGIN
END_DATA_BLOCK

DATA_BLOCK "回空结束计时"   // DB21
{ S7_Optimized_Access := 'TRUE' }
AUTHOR : Simatic
FAMILY : IEC
NAME : IEC_TMR
VERSION : 1.0
// stored: InstanceOfName IEC_TIMER
"IEC_TIMER"
BEGIN
END_DATA_BLOCK

DATA_BLOCK "慢排阀报警计时"   // DB24
{ S7_Optimized_Access := 'TRUE' }
AUTHOR : Simatic
FAMILY : IEC
NAME : IEC_TMR
VERSION : 1.0
// stored: InstanceOfName IEC_TIMER
"IEC_TIMER"
BEGIN
END_DATA_BLOCK

DATA_BLOCK "快排阀报警计时"   // DB25
{ S7_Optimized_Access := 'TRUE' }
AUTHOR : Simatic
FAMILY : IEC
NAME : IEC_TMR
VERSION : 1.0
// stored: InstanceOfName IEC_TIMER
"IEC_TIMER"
BEGIN
END_DATA_BLOCK

DATA_BLOCK "回空超时报警计时"   // DB26
{ S7_Optimized_Access := 'TRUE' }
AUTHOR : Simatic
FAMILY : IEC
NAME : IEC_TMR
VERSION : 1.0
// stored: InstanceOfName IEC_TIMER
"IEC_TIMER"
BEGIN
END_DATA_BLOCK

DATA_BLOCK "E038报警计时"   // DB29
{ S7_Optimized_Access := 'TRUE' }
AUTHOR : Simatic
FAMILY : IEC
NAME : IEC_TMR
VERSION : 1.0
// stored: InstanceOfName IEC_TIMER
"IEC_TIMER"
BEGIN
END_DATA_BLOCK

DATA_BLOCK "55℃预热复位按钮"   // DB30
{ S7_Optimized_Access := 'TRUE' }
AUTHOR : Simatic
FAMILY : IEC
NAME : IEC_TMR
VERSION : 1.0
// stored: InstanceOfName IEC_TIMER
"IEC_TIMER"
BEGIN
END_DATA_BLOCK

DATA_BLOCK "E003报警计时"   // DB31
{ S7_Optimized_Access := 'TRUE' }
AUTHOR : Simatic
FAMILY : IEC
NAME : IEC_TMR
VERSION : 1.0
// stored: InstanceOfName IEC_TIMER
"IEC_TIMER"
BEGIN
END_DATA_BLOCK

DATA_BLOCK "E004报警计时"   // DB32
{ S7_Optimized_Access := 'TRUE' }
AUTHOR : Simatic
FAMILY : IEC
NAME : IEC_TMR
VERSION : 1.0
// stored: InstanceOfName IEC_TIMER
"IEC_TIMER"
BEGIN
END_DATA_BLOCK

DATA_BLOCK "E005报警计时"   // DB33
{ S7_Optimized_Access := 'TRUE' }
AUTHOR : Simatic
FAMILY : IEC
NAME : IEC_TMR
VERSION : 1.0
// stored: InstanceOfName IEC_TIMER
"IEC_TIMER"
BEGIN
END_DATA_BLOCK

DATA_BLOCK "E006报警计时"   // DB34
{ S7_Optimized_Access := 'TRUE' }
AUTHOR : Simatic
FAMILY : IEC
NAME : IEC_TMR
VERSION : 1.0
// stored: InstanceOfName IEC_TIMER
"IEC_TIMER"
BEGIN
END_DATA_BLOCK

DATA_BLOCK "E007报警计时"   // DB35
{ S7_Optimized_Access := 'TRUE' }
AUTHOR : Simatic
FAMILY : IEC
NAME : IEC_TMR
VERSION : 1.0
// stored: InstanceOfName IEC_TIMER
"IEC_TIMER"
BEGIN
END_DATA_BLOCK

DATA_BLOCK "E008报警计时"   // DB36
{ S7_Optimized_Access := 'TRUE' }
AUTHOR : Simatic
FAMILY : IEC
NAME : IEC_TMR
VERSION : 1.0
// stored: InstanceOfName IEC_TIMER
"IEC_TIMER"
BEGIN
END_DATA_BLOCK

DATA_BLOCK "E009报警计时"   // DB37
{ S7_Optimized_Access := 'TRUE' }
AUTHOR : Simatic
FAMILY : IEC
NAME : IEC_TMR
VERSION : 1.0
// stored: InstanceOfName IEC_TIMER
"IEC_TIMER"
BEGIN
END_DATA_BLOCK

DATA_BLOCK "E013报警计时"   // DB38
{ S7_Optimized_Access := 'TRUE' }
AUTHOR : Simatic
FAMILY : IEC
NAME : IEC_TMR
VERSION : 1.0
// stored: InstanceOfName IEC_TIMER
"IEC_TIMER"
BEGIN
END_DATA_BLOCK

DATA_BLOCK "腔体加热使能计时"   // DB39
{ S7_Optimized_Access := 'TRUE' }
AUTHOR : Simatic
FAMILY : IEC
NAME : IEC_TMR
VERSION : 1.0
// stored: InstanceOfName IEC_TIMER
"IEC_TIMER"
BEGIN
END_DATA_BLOCK

DATA_BLOCK "EO16报警计时"   // DB40
{ S7_Optimized_Access := 'TRUE' }
AUTHOR : Simatic
FAMILY : IEC
NAME : IEC_TMR
VERSION : 1.0
// stored: InstanceOfName IEC_TIMER
"IEC_TIMER"
BEGIN
END_DATA_BLOCK

DATA_BLOCK "E017报警计时"   // DB41
{ S7_Optimized_Access := 'TRUE' }
AUTHOR : Simatic
FAMILY : IEC
NAME : IEC_TMR
VERSION : 1.0
// stored: InstanceOfName IEC_TIMER
"IEC_TIMER"
BEGIN
END_DATA_BLOCK

DATA_BLOCK "E018报警计时"   // DB42
{ S7_Optimized_Access := 'TRUE' }
AUTHOR : Simatic
FAMILY : IEC
NAME : IEC_TMR
VERSION : 1.0
// stored: InstanceOfName IEC_TIMER
"IEC_TIMER"
BEGIN
END_DATA_BLOCK

DATA_BLOCK "E019报警计时"   // DB43
{ S7_Optimized_Access := 'TRUE' }
AUTHOR : Simatic
FAMILY : IEC
NAME : IEC_TMR
VERSION : 1.0
// stored: InstanceOfName IEC_TIMER
"IEC_TIMER"
BEGIN
END_DATA_BLOCK

DATA_BLOCK "前门持续加热时间统计"   // DB44
{ S7_Optimized_Access := 'TRUE' }
AUTHOR : Simatic
FAMILY : IEC
NAME : CNTR
VERSION : 1.0
// stored: InstanceOfName IEC_COUNTER
"IEC_COUNTER"
BEGIN
END_DATA_BLOCK

DATA_BLOCK "后门加热持续时间统计"   // DB45
{ S7_Optimized_Access := 'TRUE' }
AUTHOR : Simatic
FAMILY : IEC
NAME : CNTR
VERSION : 1.0
// stored: InstanceOfName IEC_COUNTER
"IEC_COUNTER"
BEGIN
END_DATA_BLOCK

DATA_BLOCK "腔体后部持续加热时间统计"   // DB46
{ S7_Optimized_Access := 'TRUE' }
AUTHOR : Simatic
FAMILY : IEC
NAME : CNTR
VERSION : 1.0
// stored: InstanceOfName IEC_COUNTER
"IEC_COUNTER"
BEGIN
END_DATA_BLOCK

DATA_BLOCK "腔体前部持续加热时间统计"   // DB47
{ S7_Optimized_Access := 'TRUE' }
AUTHOR : Simatic
FAMILY : IEC
NAME : CNTR
VERSION : 1.0
// stored: InstanceOfName IEC_COUNTER
"IEC_COUNTER"
BEGIN
END_DATA_BLOCK

DATA_BLOCK "汽化器持续加热时间统计"   // DB49
{ S7_Optimized_Access := 'TRUE' }
AUTHOR : Simatic
FAMILY : IEC
NAME : CNTR
VERSION : 1.0
// stored: InstanceOfName IEC_COUNTER
"IEC_COUNTER"
BEGIN
END_DATA_BLOCK

DATA_BLOCK "E024报警计时"   // DB50
{ S7_Optimized_Access := 'TRUE' }
AUTHOR : Simatic
FAMILY : IEC
NAME : IEC_TMR
VERSION : 1.0
// stored: InstanceOfName IEC_TIMER
"IEC_TIMER"
BEGIN
END_DATA_BLOCK

DATA_BLOCK "E025报警计时"   // DB51
{ S7_Optimized_Access := 'TRUE' }
AUTHOR : Simatic
FAMILY : IEC
NAME : IEC_TMR
VERSION : 1.0
// stored: InstanceOfName IEC_TIMER
"IEC_TIMER"
BEGIN
END_DATA_BLOCK

DATA_BLOCK "E026报警计时"   // DB52
{ S7_Optimized_Access := 'TRUE' }
AUTHOR : Simatic
FAMILY : IEC
NAME : IEC_TMR
VERSION : 1.0
// stored: InstanceOfName IEC_TIMER
"IEC_TIMER"
BEGIN
END_DATA_BLOCK

DATA_BLOCK "E027报警计时"   // DB53
{ S7_Optimized_Access := 'TRUE' }
AUTHOR : Simatic
FAMILY : IEC
NAME : IEC_TMR
VERSION : 1.0
// stored: InstanceOfName IEC_TIMER
"IEC_TIMER"
BEGIN
END_DATA_BLOCK

DATA_BLOCK "E028报警计时"   // DB54
{ S7_Optimized_Access := 'TRUE' }
AUTHOR : Simatic
FAMILY : IEC
NAME : IEC_TMR
VERSION : 1.0
// stored: InstanceOfName IEC_TIMER
"IEC_TIMER"
BEGIN
END_DATA_BLOCK

DATA_BLOCK "E030报警计时"   // DB55
{ S7_Optimized_Access := 'TRUE' }
AUTHOR : Simatic
FAMILY : IEC
NAME : IEC_TMR
VERSION : 1.0
// stored: InstanceOfName IEC_TIMER
"IEC_TIMER"
BEGIN
END_DATA_BLOCK

DATA_BLOCK "E031报警计时"   // DB56
{ S7_Optimized_Access := 'TRUE' }
AUTHOR : Simatic
FAMILY : IEC
NAME : IEC_TMR
VERSION : 1.0
// stored: InstanceOfName IEC_TIMER
"IEC_TIMER"
BEGIN
END_DATA_BLOCK

DATA_BLOCK "E032报警计时"   // DB57
{ S7_Optimized_Access := 'TRUE' }
AUTHOR : Simatic
FAMILY : IEC
NAME : IEC_TMR
VERSION : 1.0
// stored: InstanceOfName IEC_TIMER
"IEC_TIMER"
BEGIN
END_DATA_BLOCK

DATA_BLOCK "E036报警计时"   // DB58
{ S7_Optimized_Access := 'TRUE' }
AUTHOR : Simatic
FAMILY : IEC
NAME : IEC_TMR
VERSION : 1.0
// stored: InstanceOfName IEC_TIMER
"IEC_TIMER"
BEGIN
END_DATA_BLOCK

DATA_BLOCK "E037报警计时"   // DB59
{ S7_Optimized_Access := 'TRUE' }
AUTHOR : Simatic
FAMILY : IEC
NAME : IEC_TMR
VERSION : 1.0
// stored: InstanceOfName IEC_TIMER
"IEC_TIMER"
BEGIN
END_DATA_BLOCK

DATA_BLOCK "报警开关复位延时"   // DB60
{ S7_Optimized_Access := 'TRUE' }
AUTHOR : Simatic
FAMILY : IEC
NAME : IEC_TMR
VERSION : 1.0
// stored: InstanceOfName IEC_TIMER
"IEC_TIMER"
BEGIN
END_DATA_BLOCK

DATA_BLOCK "保存按钮复位"   // DB61
{ S7_Optimized_Access := 'TRUE' }
AUTHOR : Simatic
FAMILY : IEC
NAME : IEC_TMR
VERSION : 1.0
// stored: InstanceOfName IEC_TIMER
"IEC_TIMER"
BEGIN
END_DATA_BLOCK

DATA_BLOCK "F010报警计时"   // DB62
{ S7_Optimized_Access := 'TRUE' }
AUTHOR : Simatic
FAMILY : IEC
NAME : IEC_TMR
VERSION : 1.0
// stored: InstanceOfName IEC_TIMER
"IEC_TIMER"
BEGIN
END_DATA_BLOCK

DATA_BLOCK "F012报警计时"   // DB63
{ S7_Optimized_Access := 'TRUE' }
AUTHOR : Simatic
FAMILY : IEC
NAME : IEC_TMR
VERSION : 1.0
// stored: InstanceOfName IEC_TIMER
"IEC_TIMER"
BEGIN
END_DATA_BLOCK

DATA_BLOCK "结束返回主菜单按钮延时"   // DB64
{ S7_Optimized_Access := 'TRUE' }
AUTHOR : Simatic
FAMILY : IEC
NAME : IEC_TMR
VERSION : 1.0
// stored: InstanceOfName IEC_TIMER
"IEC_TIMER"
BEGIN
END_DATA_BLOCK

DATA_BLOCK "E014报警计时"   // DB67
{ S7_Optimized_Access := 'TRUE' }
AUTHOR : Simatic
FAMILY : IEC
NAME : IEC_TMR
VERSION : 1.0
// stored: InstanceOfName IEC_TIMER
"IEC_TIMER"
BEGIN
END_DATA_BLOCK

DATA_BLOCK "内室负压回空延时"   // DB68
{ S7_Optimized_Access := 'TRUE' }
AUTHOR : Simatic
FAMILY : IEC
NAME : IEC_TMR
VERSION : 1.0
// stored: InstanceOfName IEC_TIMER
"IEC_TIMER"
BEGIN
END_DATA_BLOCK

DATA_BLOCK "运行时页面强制跳转"   // DB69
{ S7_Optimized_Access := 'TRUE' }
AUTHOR : Simatic
FAMILY : IEC
NAME : IEC_TMR
VERSION : 1.0
// stored: InstanceOfName IEC_TIMER
"IEC_TIMER"
BEGIN
END_DATA_BLOCK

DATA_BLOCK "启动按钮复位"   // DB72
{ S7_Optimized_Access := 'TRUE' }
AUTHOR : Simatic
FAMILY : IEC
NAME : IEC_TMR
VERSION : 1.0
// stored: InstanceOfName IEC_TIMER
"IEC_TIMER"
BEGIN
END_DATA_BLOCK

DATA_BLOCK "设备维护复位按钮"   // DB73
{ S7_Optimized_Access := 'TRUE' }
AUTHOR : Simatic
FAMILY : IEC
NAME : IEC_TMR
VERSION : 1.0
// stored: InstanceOfName IEC_TIMER
"IEC_TIMER"
BEGIN
END_DATA_BLOCK

DATA_BLOCK "报警计时"   // DB75
{ S7_Optimized_Access := 'TRUE' }
AUTHOR : Simatic
FAMILY : IEC
NAME : IEC_TMR
VERSION : 1.0
// stored: InstanceOfName IEC_TIMER
"IEC_TIMER"
BEGIN
END_DATA_BLOCK

DATA_BLOCK "报警确认按钮复位计时"   // DB78
{ S7_Optimized_Access := 'TRUE' }
AUTHOR : Simatic
FAMILY : IEC
NAME : IEC_TMR
VERSION : 1.0
// stored: InstanceOfName IEC_TIMER
"IEC_TIMER"
BEGIN
END_DATA_BLOCK

DATA_BLOCK "数据传递按钮复位"   // DB79
{ S7_Optimized_Access := 'TRUE' }
AUTHOR : Simatic
FAMILY : IEC
NAME : IEC_TMR
VERSION : 1.0
// stored: InstanceOfName IEC_TIMER
"IEC_TIMER"
BEGIN
END_DATA_BLOCK

DATA_BLOCK "催化箱加热时间统计"   // DB80
{ S7_Optimized_Access := 'TRUE' }
AUTHOR : Simatic
FAMILY : IEC
NAME : CNTR
VERSION : 1.0
// stored: InstanceOfName IEC_COUNTER
"IEC_COUNTER"
BEGIN
END_DATA_BLOCK

DATA_BLOCK "阶段跳转延时"   // DB81
{ S7_Optimized_Access := 'TRUE' }
AUTHOR : Simatic
FAMILY : IEC
NAME : IEC_TMR
VERSION : 1.0
// stored: InstanceOfName IEC_TIMER
"IEC_TIMER"
BEGIN
END_DATA_BLOCK

DATA_BLOCK "加湿阶段跳转延时"   // DB82
{ S7_Optimized_Access := 'TRUE' }
AUTHOR : Simatic
FAMILY : IEC
NAME : IEC_TMR
VERSION : 1.0
// stored: InstanceOfName IEC_TIMER
"IEC_TIMER"
BEGIN
END_DATA_BLOCK

DATA_BLOCK "结束跳转阶段延时"   // DB83
{ S7_Optimized_Access := 'TRUE' }
AUTHOR : Simatic
FAMILY : IEC
NAME : IEC_TMR
VERSION : 1.0
// stored: InstanceOfName IEC_TIMER
"IEC_TIMER"
BEGIN
END_DATA_BLOCK

DATA_BLOCK "运行时间统计"   // DB86
{ S7_Optimized_Access := 'TRUE' }
AUTHOR : Simatic
FAMILY : IEC
NAME : IEC_TMR
VERSION : 1.0
// stored: InstanceOfName IEC_TIMER
"IEC_TIMER"
BEGIN
END_DATA_BLOCK

DATA_BLOCK "正常结束标志复位"   // DB90
{ S7_Optimized_Access := 'TRUE' }
AUTHOR : Simatic
FAMILY : IEC
NAME : IEC_TMR
VERSION : 1.0
// stored: InstanceOfName IEC_TIMER
"IEC_TIMER"
BEGIN
END_DATA_BLOCK

DATA_BLOCK "催化剂维护按钮复位"   // DB92
{ S7_Optimized_Access := 'TRUE' }
AUTHOR : Simatic
FAMILY : IEC
NAME : IEC_TMR
VERSION : 1.0
// stored: InstanceOfName IEC_TIMER
"IEC_TIMER"
BEGIN
END_DATA_BLOCK

DATA_BLOCK "开前门按钮复位"   // DB93
{ S7_Optimized_Access := 'TRUE' }
AUTHOR : Simatic
FAMILY : IEC
NAME : IEC_TMR
VERSION : 1.0
// stored: InstanceOfName IEC_TIMER
"IEC_TIMER"
BEGIN
END_DATA_BLOCK

DATA_BLOCK "关前门按钮复位"   // DB94
{ S7_Optimized_Access := 'TRUE' }
AUTHOR : Simatic
FAMILY : IEC
NAME : IEC_TMR
VERSION : 1.0
// stored: InstanceOfName IEC_TIMER
"IEC_TIMER"
BEGIN
END_DATA_BLOCK

DATA_BLOCK "开后门按钮复位"   // DB95
{ S7_Optimized_Access := 'TRUE' }
AUTHOR : Simatic
FAMILY : IEC
NAME : IEC_TMR
VERSION : 1.0
// stored: InstanceOfName IEC_TIMER
"IEC_TIMER"
BEGIN
END_DATA_BLOCK

DATA_BLOCK "关后门按钮复位"   // DB96
{ S7_Optimized_Access := 'TRUE' }
AUTHOR : Simatic
FAMILY : IEC
NAME : IEC_TMR
VERSION : 1.0
// stored: InstanceOfName IEC_TIMER
"IEC_TIMER"
BEGIN
END_DATA_BLOCK

DATA_BLOCK "新报警标识复位计时"   // DB98
{ S7_Optimized_Access := 'TRUE' }
AUTHOR : Simatic
FAMILY : IEC
NAME : IEC_TMR
VERSION : 1.0
// stored: InstanceOfName IEC_TIMER
"IEC_TIMER"
BEGIN
END_DATA_BLOCK

DATA_BLOCK "进入预热页面延时"   // DB101
{ S7_Optimized_Access := 'TRUE' }
AUTHOR : Simatic
FAMILY : IEC
NAME : IEC_TMR
VERSION : 1.0
// stored: InstanceOfName IEC_TIMER
"IEC_TIMER"
BEGIN
END_DATA_BLOCK

DATA_BLOCK "加湿湿度达到设定湿度延时"   // DB105
{ S7_Optimized_Access := 'TRUE' }
AUTHOR : Simatic
FAMILY : IEC
NAME : IEC_TMR
VERSION : 1.0
// stored: InstanceOfName IEC_TIMER
"IEC_TIMER"
BEGIN
END_DATA_BLOCK

DATA_BLOCK "灭菌报表打印时间间隔"   // DB106
{ S7_Optimized_Access := 'TRUE' }
AUTHOR : Simatic
FAMILY : IEC
NAME : IEC_TMR
VERSION : 1.0
// stored: InstanceOfName IEC_TIMER
"IEC_TIMER"
BEGIN
END_DATA_BLOCK

DATA_BLOCK "保压正常结束清零延时"   // DB107
{ S7_Optimized_Access := 'TRUE' }
AUTHOR : Simatic
FAMILY : IEC
NAME : IEC_TMR
VERSION : 1.0
// stored: InstanceOfName IEC_TIMER
"IEC_TIMER"
BEGIN
END_DATA_BLOCK

DATA_BLOCK "恢复默认按钮复位"   // DB108
{ S7_Optimized_Access := 'TRUE' }
AUTHOR : Simatic
FAMILY : IEC
NAME : IEC_TMR
VERSION : 1.0
// stored: InstanceOfName IEC_TIMER
"IEC_TIMER"
BEGIN
END_DATA_BLOCK

DATA_BLOCK "E029报警延时"   // DB113
{ S7_Optimized_Access := 'TRUE' }
AUTHOR : Simatic
FAMILY : IEC
NAME : IEC_TMR
VERSION : 1.0
// stored: InstanceOfName IEC_TIMER
"IEC_TIMER"
BEGIN
END_DATA_BLOCK

DATA_BLOCK "灭菌压力过高报警延时"   // DB114
{ S7_Optimized_Access := 'TRUE' }
AUTHOR : Simatic
FAMILY : IEC
NAME : IEC_TMR
VERSION : 1.0
// stored: InstanceOfName IEC_TIMER
"IEC_TIMER"
BEGIN
END_DATA_BLOCK

DATA_BLOCK "保压异常结束运行标志延时"   // DB115
{ S7_Optimized_Access := 'TRUE' }
AUTHOR : Simatic
FAMILY : IEC
NAME : IEC_TMR
VERSION : 1.0
// stored: InstanceOfName IEC_TIMER
"IEC_TIMER"
BEGIN
END_DATA_BLOCK

DATA_BLOCK "时钟冻结延时"   // DB116
{ S7_Optimized_Access := 'TRUE' }
AUTHOR : Simatic
FAMILY : IEC
NAME : IEC_TMR
VERSION : 1.0
// stored: InstanceOfName IEC_TIMER
"IEC_TIMER"
BEGIN
END_DATA_BLOCK

DATA_BLOCK "通风回空阀开启延时"   // DB117
{ S7_Optimized_Access := 'TRUE' }
AUTHOR : Simatic
FAMILY : IEC
NAME : IEC_TMR
VERSION : 1.0
// stored: InstanceOfName IEC_TIMER
"IEC_TIMER"
BEGIN
END_DATA_BLOCK

DATA_BLOCK "E012报警延时"   // DB118
{ S7_Optimized_Access := 'TRUE' }
AUTHOR : Simatic
FAMILY : IEC
NAME : IEC_TMR
VERSION : 1.0
// stored: InstanceOfName IEC_TIMER
"IEC_TIMER"
BEGIN
END_DATA_BLOCK

DATA_BLOCK "E010报警延时"   // DB119
{ S7_Optimized_Access := 'TRUE' }
AUTHOR : Simatic
FAMILY : IEC
NAME : IEC_TMR
VERSION : 1.0
// stored: InstanceOfName IEC_TIMER
"IEC_TIMER"
BEGIN
END_DATA_BLOCK

DATA_BLOCK "加湿阶段回空延时"   // DB120
{ S7_Optimized_Access := 'TRUE' }
AUTHOR : Simatic
FAMILY : IEC
NAME : IEC_TMR
VERSION : 1.0
// stored: InstanceOfName IEC_TIMER
"IEC_TIMER"
BEGIN
END_DATA_BLOCK

DATA_BLOCK "防页面卡倒计时页面"   // DB121
{ S7_Optimized_Access := 'TRUE' }
AUTHOR : Simatic
FAMILY : IEC
NAME : IEC_TMR
VERSION : 1.0
// stored: InstanceOfName IEC_TIMER
"IEC_TIMER"
BEGIN
END_DATA_BLOCK

DATA_BLOCK "E015报警计时"   // DB122
{ S7_Optimized_Access := 'TRUE' }
AUTHOR : Simatic
FAMILY : IEC
NAME : IEC_TMR
VERSION : 1.0
// stored: InstanceOfName IEC_TIMER
"IEC_TIMER"
BEGIN
END_DATA_BLOCK

DATA_BLOCK "强制恢复默认IP延时"   // DB123
{ S7_Optimized_Access := 'TRUE' }
AUTHOR : Simatic
FAMILY : IEC
NAME : IEC_TMR
VERSION : 1.0
// stored: InstanceOfName IEC_TIMER
"IEC_TIMER"
BEGIN
END_DATA_BLOCK

DATA_BLOCK "手动退出按钮复位"   // DB124
{ S7_Optimized_Access := 'TRUE' }
AUTHOR : Simatic
FAMILY : IEC
NAME : IEC_TMR
VERSION : 1.0
// stored: InstanceOfName IEC_TIMER
"IEC_TIMER"
BEGIN
END_DATA_BLOCK

DATA_BLOCK "通风快抽空阀开启延时"   // DB125
{ S7_Optimized_Access := 'TRUE' }
AUTHOR : Simatic
FAMILY : IEC
NAME : IEC_TMR
VERSION : 1.0
// stored: InstanceOfName IEC_TIMER
"IEC_TIMER"
BEGIN
END_DATA_BLOCK

DATA_BLOCK "湿度报警延时"   // DB126
{ S7_Optimized_Access := 'TRUE' }
AUTHOR : Simatic
FAMILY : IEC
NAME : IEC_TMR
VERSION : 1.0
// stored: InstanceOfName IEC_TIMER
"IEC_TIMER"
BEGIN
END_DATA_BLOCK

DATA_BLOCK "穿刺初不记录压力值"   // DB127
{ S7_Optimized_Access := 'TRUE' }
AUTHOR : Simatic
FAMILY : IEC
NAME : IEC_TMR
VERSION : 1.0
// stored: InstanceOfName IEC_TIMER
"IEC_TIMER"
BEGIN
END_DATA_BLOCK

DATA_BLOCK "急停报警延时"   // DB130
{ S7_Optimized_Access := 'TRUE' }
AUTHOR : Simatic
FAMILY : IEC
NAME : IEC_TMR
VERSION : 1.0
// stored: InstanceOfName IEC_TIMER
"IEC_TIMER"
BEGIN
END_DATA_BLOCK

DATA_BLOCK "E022报警延时"   // DB131
{ S7_Optimized_Access := 'TRUE' }
AUTHOR : Simatic
FAMILY : IEC
NAME : IEC_TMR
VERSION : 1.0
// stored: InstanceOfName IEC_TIMER
"IEC_TIMER"
BEGIN
END_DATA_BLOCK

DATA_BLOCK "E023报警延时"   // DB132
{ S7_Optimized_Access := 'TRUE' }
AUTHOR : Simatic
FAMILY : IEC
NAME : IEC_TMR
VERSION : 1.0
// stored: InstanceOfName IEC_TIMER
"IEC_TIMER"
BEGIN
END_DATA_BLOCK

DATA_BLOCK "运行标志延时复位"   // DB133
{ S7_Optimized_Access := 'TRUE' }
AUTHOR : Simatic
FAMILY : IEC
NAME : IEC_TMR
VERSION : 1.0
// stored: InstanceOfName IEC_TIMER
"IEC_TIMER"
BEGIN
END_DATA_BLOCK

DATA_BLOCK "运行标志延时复位1"   // DB134
{ S7_Optimized_Access := 'TRUE' }
AUTHOR : Simatic
FAMILY : IEC
NAME : IEC_TMR
VERSION : 1.0
// stored: InstanceOfName IEC_TIMER
"IEC_TIMER"
BEGIN
END_DATA_BLOCK

DATA_BLOCK "上电时间统计定时器"   // DB135
{ S7_Optimized_Access := 'TRUE' }
AUTHOR : Simatic
FAMILY : IEC
NAME : IEC_TMR
VERSION : 1.0
// stored: InstanceOfName IEC_TIMER
"IEC_TIMER"
BEGIN
END_DATA_BLOCK

DATA_BLOCK "程序结束后计时"   // DB137
{ S7_Optimized_Access := 'TRUE' }
AUTHOR : Simatic
FAMILY : IEC
NAME : IEC_TMR
VERSION : 1.0
// stored: InstanceOfName IEC_TIMER
"IEC_TIMER"
BEGIN
END_DATA_BLOCK

DATA_BLOCK "达到开门条件延时十秒"   // DB138
{ S7_Optimized_Access := 'TRUE' }
AUTHOR : Simatic
FAMILY : IEC
NAME : IEC_TMR
VERSION : 1.0
// stored: InstanceOfName IEC_TIMER
"IEC_TIMER"
BEGIN
END_DATA_BLOCK

DATA_BLOCK "回空等待5分钟计时器"   // DB139
{ S7_Optimized_Access := 'TRUE' }
AUTHOR : Simatic
FAMILY : IEC
NAME : IEC_TMR
VERSION : 1.0
// stored: InstanceOfName IEC_TIMER
"IEC_TIMER"
BEGIN
END_DATA_BLOCK

DATA_BLOCK "脉动抽空运行时间"   // DB140
{ S7_Optimized_Access := 'TRUE' }
AUTHOR : Simatic
FAMILY : IEC
NAME : IEC_TMR
VERSION : 1.0
// stored: InstanceOfName IEC_TIMER
"IEC_TIMER"
BEGIN
END_DATA_BLOCK

DATA_BLOCK "脉动回空运行时间"   // DB141
{ S7_Optimized_Access := 'TRUE' }
AUTHOR : Simatic
FAMILY : IEC
NAME : IEC_TMR
VERSION : 1.0
// stored: InstanceOfName IEC_TIMER
"IEC_TIMER"
BEGIN
END_DATA_BLOCK

DATA_BLOCK "穿刺初不记录压力值2"   // DB144
{ S7_Optimized_Access := 'TRUE' }
AUTHOR : Simatic
FAMILY : IEC
NAME : IEC_TMR
VERSION : 1.0
// stored: InstanceOfName IEC_TIMER
"IEC_TIMER"
BEGIN
END_DATA_BLOCK

DATA_BLOCK "EO011报警延时"   // DB146
{ S7_Optimized_Access := 'TRUE' }
AUTHOR : Simatic
FAMILY : IEC
NAME : IEC_TMR
VERSION : 1.0
// stored: InstanceOfName IEC_TIMER
"IEC_TIMER"
BEGIN
END_DATA_BLOCK

DATA_BLOCK "双泵切换标志清零延时"   // DB147
{ S7_Optimized_Access := 'TRUE' }
AUTHOR : Simatic
FAMILY : IEC
NAME : IEC_TMR
VERSION : 1.0
// stored: InstanceOfName IEC_TIMER
"IEC_TIMER"
BEGIN
END_DATA_BLOCK

DATA_BLOCK "预热报表打印间隔"   // DB152
{ S7_Optimized_Access := 'TRUE' }
AUTHOR : Simatic
FAMILY : IEC
NAME : IEC_TMR
VERSION : 1.0
// stored: InstanceOfName IEC_TIMER
"IEC_TIMER"
BEGIN
END_DATA_BLOCK

DATA_BLOCK "通风报表打印间隔"   // DB153
{ S7_Optimized_Access := 'TRUE' }
AUTHOR : Simatic
FAMILY : IEC
NAME : IEC_TMR
VERSION : 1.0
// stored: InstanceOfName IEC_TIMER
"IEC_TIMER"
BEGIN
END_DATA_BLOCK

DATA_BLOCK "强制恢复IP复位"   // DB154
{ S7_Optimized_Access := 'TRUE' }
AUTHOR : Simatic
FAMILY : IEC
NAME : IEC_TMR
VERSION : 1.0
// stored: InstanceOfName IEC_TIMER
"IEC_TIMER"
BEGIN
END_DATA_BLOCK

DATA_BLOCK "灭菌时间统计"   // DB155
{ S7_Optimized_Access := 'TRUE' }
AUTHOR : Simatic
FAMILY : IEC
NAME : IEC_TMR
VERSION : 1.0
// stored: InstanceOfName IEC_TIMER
"IEC_TIMER"
BEGIN
END_DATA_BLOCK

DATA_BLOCK "保压报表打印间隔"   // DB156
{ S7_Optimized_Access := 'TRUE' }
AUTHOR : Simatic
FAMILY : IEC
NAME : IEC_TMR
VERSION : 1.0
// stored: InstanceOfName IEC_TIMER
"IEC_TIMER"
BEGIN
END_DATA_BLOCK

DATA_BLOCK "加湿报表打印间隔"   // DB157
{ S7_Optimized_Access := 'TRUE' }
AUTHOR : Simatic
FAMILY : IEC
NAME : IEC_TMR
VERSION : 1.0
// stored: InstanceOfName IEC_TIMER
"IEC_TIMER"
BEGIN
END_DATA_BLOCK

DATA_BLOCK "加药报表打印间隔"   // DB158
{ S7_Optimized_Access := 'TRUE' }
AUTHOR : Simatic
FAMILY : IEC
NAME : IEC_TMR
VERSION : 1.0
// stored: InstanceOfName IEC_TIMER
"IEC_TIMER"
BEGIN
END_DATA_BLOCK

DATA_BLOCK "预处理小阶段时间统计"   // DB159
{ S7_Optimized_Access := 'TRUE' }
AUTHOR : Simatic
FAMILY : IEC
NAME : IEC_TMR
VERSION : 1.0
// stored: InstanceOfName IEC_TIMER
"IEC_TIMER"
BEGIN
END_DATA_BLOCK

DATA_BLOCK "脉动报表打印间隔"   // DB163
{ S7_Optimized_Access := 'TRUE' }
AUTHOR : Simatic
FAMILY : IEC
NAME : IEC_TMR
VERSION : 1.0
// stored: InstanceOfName IEC_TIMER
"IEC_TIMER"
BEGIN
END_DATA_BLOCK

DATA_BLOCK "结束报表打印间隔"   // DB164
{ S7_Optimized_Access := 'TRUE' }
AUTHOR : Simatic
FAMILY : IEC
NAME : IEC_TMR
VERSION : 1.0
// stored: InstanceOfName IEC_TIMER
"IEC_TIMER"
BEGIN
END_DATA_BLOCK

DATA_BLOCK "保压小阶段时间统计"   // DB165
{ S7_Optimized_Access := 'TRUE' }
AUTHOR : Simatic
FAMILY : IEC
NAME : IEC_TMR
VERSION : 1.0
// stored: InstanceOfName IEC_TIMER
"IEC_TIMER"
BEGIN
END_DATA_BLOCK

DATA_BLOCK "加湿大阶段时间统计"   // DB166
{ S7_Optimized_Access := 'TRUE' }
AUTHOR : Simatic
FAMILY : IEC
NAME : IEC_TMR
VERSION : 1.0
// stored: InstanceOfName IEC_TIMER
"IEC_TIMER"
BEGIN
END_DATA_BLOCK

DATA_BLOCK "加湿小阶段时间统计"   // DB167
{ S7_Optimized_Access := 'TRUE' }
AUTHOR : Simatic
FAMILY : IEC
NAME : IEC_TMR
VERSION : 1.0
// stored: InstanceOfName IEC_TIMER
"IEC_TIMER"
BEGIN
END_DATA_BLOCK

DATA_BLOCK "加药大阶段时间统计"   // DB168
{ S7_Optimized_Access := 'TRUE' }
AUTHOR : Simatic
FAMILY : IEC
NAME : IEC_TMR
VERSION : 1.0
// stored: InstanceOfName IEC_TIMER
"IEC_TIMER"
BEGIN
END_DATA_BLOCK

DATA_BLOCK "加药小阶段时间统计"   // DB169
{ S7_Optimized_Access := 'TRUE' }
AUTHOR : Simatic
FAMILY : IEC
NAME : IEC_TMR
VERSION : 1.0
// stored: InstanceOfName IEC_TIMER
"IEC_TIMER"
BEGIN
END_DATA_BLOCK

DATA_BLOCK "脉动大阶段时间统计"   // DB170
{ S7_Optimized_Access := 'TRUE' }
AUTHOR : Simatic
FAMILY : IEC
NAME : IEC_TMR
VERSION : 1.0
// stored: InstanceOfName IEC_TIMER
"IEC_TIMER"
BEGIN
END_DATA_BLOCK

DATA_BLOCK "脉动小阶段时间统计"   // DB171
{ S7_Optimized_Access := 'TRUE' }
AUTHOR : Simatic
FAMILY : IEC
NAME : IEC_TMR
VERSION : 1.0
// stored: InstanceOfName IEC_TIMER
"IEC_TIMER"
BEGIN
END_DATA_BLOCK

DATA_BLOCK "通风大阶段时间统计"   // DB172
{ S7_Optimized_Access := 'TRUE' }
AUTHOR : Simatic
FAMILY : IEC
NAME : IEC_TMR
VERSION : 1.0
// stored: InstanceOfName IEC_TIMER
"IEC_TIMER"
BEGIN
END_DATA_BLOCK

DATA_BLOCK "通风小阶段时间统计"   // DB173
{ S7_Optimized_Access := 'TRUE' }
AUTHOR : Simatic
FAMILY : IEC
NAME : IEC_TMR
VERSION : 1.0
// stored: InstanceOfName IEC_TIMER
"IEC_TIMER"
BEGIN
END_DATA_BLOCK

DATA_BLOCK "保压异常结束大阶段清零"   // DB174
{ S7_Optimized_Access := 'TRUE' }
AUTHOR : Simatic
FAMILY : IEC
NAME : IEC_TMR
VERSION : 1.0
// stored: InstanceOfName IEC_TIMER
"IEC_TIMER"
BEGIN
END_DATA_BLOCK

DATA_BLOCK "结束大阶段时间统计"   // DB175
{ S7_Optimized_Access := 'TRUE' }
AUTHOR : Simatic
FAMILY : IEC
NAME : IEC_TMR
VERSION : 1.0
// stored: InstanceOfName IEC_TIMER
"IEC_TIMER"
BEGIN
END_DATA_BLOCK

DATA_BLOCK "结束小阶段时间统计"   // DB176
{ S7_Optimized_Access := 'TRUE' }
AUTHOR : Simatic
FAMILY : IEC
NAME : IEC_TMR
VERSION : 1.0
// stored: InstanceOfName IEC_TIMER
"IEC_TIMER"
BEGIN
END_DATA_BLOCK

DATA_BLOCK "紧急脉动大阶段时间统计"   // DB177
{ S7_Optimized_Access := 'TRUE' }
AUTHOR : Simatic
FAMILY : IEC
NAME : IEC_TMR
VERSION : 1.0
// stored: InstanceOfName IEC_TIMER
"IEC_TIMER"
BEGIN
END_DATA_BLOCK

DATA_BLOCK "紧急脉动小阶段时间统计"   // DB178
{ S7_Optimized_Access := 'TRUE' }
AUTHOR : Simatic
FAMILY : IEC
NAME : IEC_TMR
VERSION : 1.0
// stored: InstanceOfName IEC_TIMER
"IEC_TIMER"
BEGIN
END_DATA_BLOCK

DATA_BLOCK "紧急通风大阶段时间统计"   // DB179
{ S7_Optimized_Access := 'TRUE' }
AUTHOR : Simatic
FAMILY : IEC
NAME : IEC_TMR
VERSION : 1.0
// stored: InstanceOfName IEC_TIMER
"IEC_TIMER"
BEGIN
END_DATA_BLOCK

DATA_BLOCK "紧急通风小阶段时间统计"   // DB180
{ S7_Optimized_Access := 'TRUE' }
AUTHOR : Simatic
FAMILY : IEC
NAME : IEC_TMR
VERSION : 1.0
// stored: InstanceOfName IEC_TIMER
"IEC_TIMER"
BEGIN
END_DATA_BLOCK

DATA_BLOCK "紧急标志清零延时"   // DB181
{ S7_Optimized_Access := 'TRUE' }
AUTHOR : Simatic
FAMILY : IEC
NAME : IEC_TMR
VERSION : 1.0
// stored: InstanceOfName IEC_TIMER
"IEC_TIMER"
BEGIN
END_DATA_BLOCK

DATA_BLOCK "结束后大阶段强制复位延时"   // DB182
{ S7_Optimized_Access := 'TRUE' }
AUTHOR : Simatic
FAMILY : IEC
NAME : IEC_TMR
VERSION : 1.0
// stored: InstanceOfName IEC_TIMER
"IEC_TIMER"
BEGIN
END_DATA_BLOCK

DATA_BLOCK "内室压力低于250mbar滤波"   // DB183
{ S7_Optimized_Access := 'TRUE' }
AUTHOR : Simatic
FAMILY : IEC
NAME : IEC_TMR
VERSION : 1.0
// stored: InstanceOfName IEC_TIMER
"IEC_TIMER"
BEGIN
END_DATA_BLOCK

DATA_BLOCK "网络设置按钮复位"   // DB1001
{ S7_Optimized_Access := 'TRUE' }
AUTHOR : Simatic
FAMILY : IEC
NAME : IEC_TMR
VERSION : 1.0
// stored: InstanceOfName IEC_TIMER
"IEC_TIMER"
BEGIN
END_DATA_BLOCK

// folder: (top level)

ORGANIZATION_BLOCK "Startup"   // OB100, LAD, Startup
TITLE = "Complete Restart"
{ S7_Optimized_Access := 'TRUE' }
VERSION : 0.1
   VAR_INPUT
      LostRetentive : Bool;   // True if retentive data are lost
      LostRTC : Bool;   // True if date and time are lost
   END_VAR
   VAR_TEMP
      BUSY1 : Bool;
      BUSY2 : Bool;
      BUSY3 : Bool;
   END_VAR
BEGIN

REGION Network 1: 单扉
   // "触摸屏".设备配置.%X5   为0时 为单扉   为1时为双扉
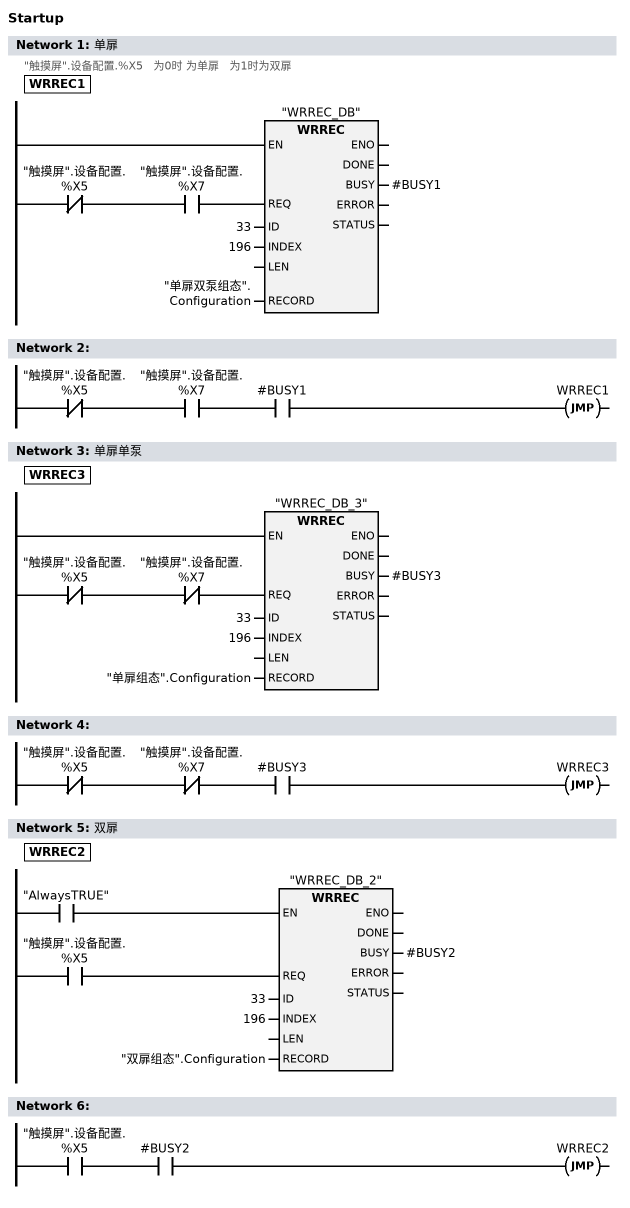
   WRREC1:
   "WRREC_DB"(REQ := NOT "触摸屏".设备配置.%X5 AND "触摸屏".设备配置.%X7,   // WRREC
              ID := 33,
              INDEX := 196,
              RECORD := "单扉双泵组态".Configuration,
              BUSY => #BUSY1);
END_REGION

REGION Network 2
   RUNG wire#powerrail
      I_Contact( "触摸屏".设备配置.%X5 )
      Contact( "触摸屏".设备配置.%X7 )
      Contact( #BUSY1 )
      JumpCoil( WRREC1 )
   END_RUNG
   // the same network as SCL:
   IF NOT "触摸屏".设备配置.%X5 AND "触摸屏".设备配置.%X7 AND #BUSY1 THEN GOTO WRREC1; END_IF;
END_REGION

REGION Network 3: 单扉单泵
   WRREC3:
   "WRREC_DB_3"(REQ := NOT "触摸屏".设备配置.%X5 AND NOT "触摸屏".设备配置.%X7,   // WRREC
                ID := 33,
                INDEX := 196,
                RECORD := "单扉组态".Configuration,
                BUSY => #BUSY3);
END_REGION

REGION Network 4
   RUNG wire#powerrail
      I_Contact( "触摸屏".设备配置.%X5 )
      I_Contact( "触摸屏".设备配置.%X7 )
      Contact( #BUSY3 )
      JumpCoil( WRREC3 )
   END_RUNG
   // the same network as SCL:
   IF NOT "触摸屏".设备配置.%X5 AND NOT "触摸屏".设备配置.%X7 AND #BUSY3 THEN GOTO WRREC3; END_IF;
END_REGION

REGION Network 5: 双扉
   WRREC2:
   IF "AlwaysTRUE" THEN
       "WRREC_DB_2"(REQ := "触摸屏".设备配置.%X5, ID := 33, INDEX := 196, RECORD := "双扉组态".Configuration, BUSY => #BUSY2);   // WRREC
   END_IF;
END_REGION

REGION Network 6
   RUNG wire#powerrail
      Contact( "触摸屏".设备配置.%X5 )
      Contact( #BUSY2 )
      JumpCoil( WRREC2 )
   END_RUNG
   // the same network as SCL:
   IF "触摸屏".设备配置.%X5 AND #BUSY2 THEN GOTO WRREC2; END_IF;
END_REGION
END_ORGANIZATION_BLOCK

// folder: 1 初始化+版本

FUNCTION "初始化＋版本号" : Void   // FC1, LAD
{ S7_Optimized_Access := 'TRUE' }
VERSION : 0.1
// EO3000-N260610 修复保压测试程序温度问题,预热温度显示
// EO3000-N260909 增加韩语打印 PLC仅变更版本后 其余程序没变化
BEGIN

REGION Network 1: 程序版本号
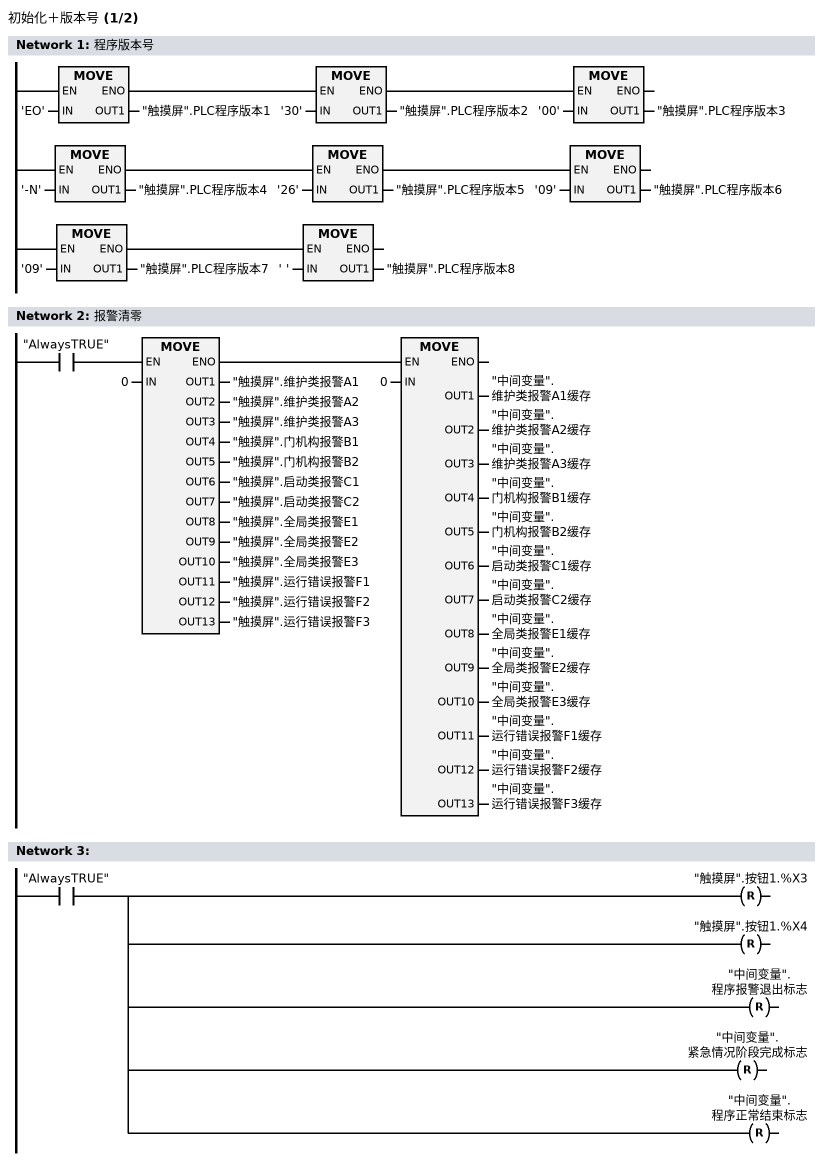
   RUNG wire#powerrail
      Move(in := 'EO', out1 => "触摸屏".PLC程序版本1)
      Move(in := '30', out1 => "触摸屏".PLC程序版本2)
      Move(in := '00', out1 => "触摸屏".PLC程序版本3)
   END_RUNG
   RUNG wire#powerrail
      Move(in := '-N', out1 => "触摸屏".PLC程序版本4)
      Move(in := '26', out1 => "触摸屏".PLC程序版本5)
      Move(in := '09', out1 => "触摸屏".PLC程序版本6)
   END_RUNG
   RUNG wire#powerrail
      Move(in := '09', out1 => "触摸屏".PLC程序版本7)
      Move(in := ' ', out1 => "触摸屏".PLC程序版本8)
   END_RUNG
   // the same network as SCL:
   "触摸屏".PLC程序版本1 := 'EO';
   "触摸屏".PLC程序版本2 := '30';
   "触摸屏".PLC程序版本3 := '00';
   "触摸屏".PLC程序版本4 := '-N';
   "触摸屏".PLC程序版本5 := '26';
   "触摸屏".PLC程序版本6 := '09';
   "触摸屏".PLC程序版本7 := '09';
   "触摸屏".PLC程序版本8 := ' ';
END_REGION

REGION Network 2: 报警清零
   RUNG wire#powerrail
      Contact( "AlwaysTRUE" )
      Move(in := 0, out1 => "触摸屏".维护类报警A1, out2 => "触摸屏".维护类报警A2, out3 => "触摸屏".维护类报警A3, out4 => "触摸屏".门机构报警B1, out5 => "触摸屏".门机构报警B2, out6 => "触摸屏".启动类报警C1, out7 => "触摸屏".启动类报警C2, out8 => "触摸屏".全局类报警E1, out9 => "触摸屏".全局类报警E2, out10 => "触摸屏".全局类报警E3, out11 => "触摸屏".运行错误报警F1, out12 => "触摸屏".运行错误报警F2, out13 => "触摸屏".运行错误报警F3)
      Move(in := 0, out1 => "中间变量".维护类报警A1缓存, out2 => "中间变量".维护类报警A2缓存, out3 => "中间变量".维护类报警A3缓存, out4 => "中间变量".门机构报警B1缓存, out5 => "中间变量".门机构报警B2缓存, out6 => "中间变量".启动类报警C1缓存, out7 => "中间变量".启动类报警C2缓存, out8 => "中间变量".全局类报警E1缓存, out9 => "中间变量".全局类报警E2缓存, out10 => "中间变量".全局类报警E3缓存, out11 => "中间变量".运行错误报警F1缓存, out12 => "中间变量".运行错误报警F2缓存, out13 => "中间变量".运行错误报警F3缓存)
   END_RUNG
   // the same network as SCL:
   IF "AlwaysTRUE" THEN
       "触摸屏".维护类报警A1 := 0;
       "触摸屏".维护类报警A2 := 0;
       "触摸屏".维护类报警A3 := 0;
       "触摸屏".门机构报警B1 := 0;
       "触摸屏".门机构报警B2 := 0;
       "触摸屏".启动类报警C1 := 0;
       "触摸屏".启动类报警C2 := 0;
       "触摸屏".全局类报警E1 := 0;
       "触摸屏".全局类报警E2 := 0;
       "触摸屏".全局类报警E3 := 0;
       "触摸屏".运行错误报警F1 := 0;
       "触摸屏".运行错误报警F2 := 0;
       "触摸屏".运行错误报警F3 := 0;
       "中间变量".维护类报警A1缓存 := 0;
       "中间变量".维护类报警A2缓存 := 0;
       "中间变量".维护类报警A3缓存 := 0;
       "中间变量".门机构报警B1缓存 := 0;
       "中间变量".门机构报警B2缓存 := 0;
       "中间变量".启动类报警C1缓存 := 0;
       "中间变量".启动类报警C2缓存 := 0;
       "中间变量".全局类报警E1缓存 := 0;
       "中间变量".全局类报警E2缓存 := 0;
       "中间变量".全局类报警E3缓存 := 0;
       "中间变量".运行错误报警F1缓存 := 0;
       "中间变量".运行错误报警F2缓存 := 0;
       "中间变量".运行错误报警F3缓存 := 0;
   END_IF;
END_REGION

REGION Network 3
   RUNG wire#powerrail
      Contact( "AlwaysTRUE" )
      wire#w1
      R_Coil( "触摸屏".按钮1.%X3 )
   END_RUNG
   RUNG wire#w1
      R_Coil( "触摸屏".按钮1.%X4 )
   END_RUNG
   RUNG wire#w1
      R_Coil( "中间变量".程序报警退出标志 )
   END_RUNG
   RUNG wire#w1
      R_Coil( "中间变量".紧急情况阶段完成标志 )
   END_RUNG
   RUNG wire#w1
      R_Coil( "中间变量".程序正常结束标志 )
   END_RUNG
   // the same network as SCL:
   IF "AlwaysTRUE" THEN
       "触摸屏".按钮1.%X3 := FALSE;
       "触摸屏".按钮1.%X4 := FALSE;
       "中间变量".程序报警退出标志 := FALSE;
       "中间变量".紧急情况阶段完成标志 := FALSE;
       "中间变量".程序正常结束标志 := FALSE;
   END_IF;
END_REGION

REGION Network 4
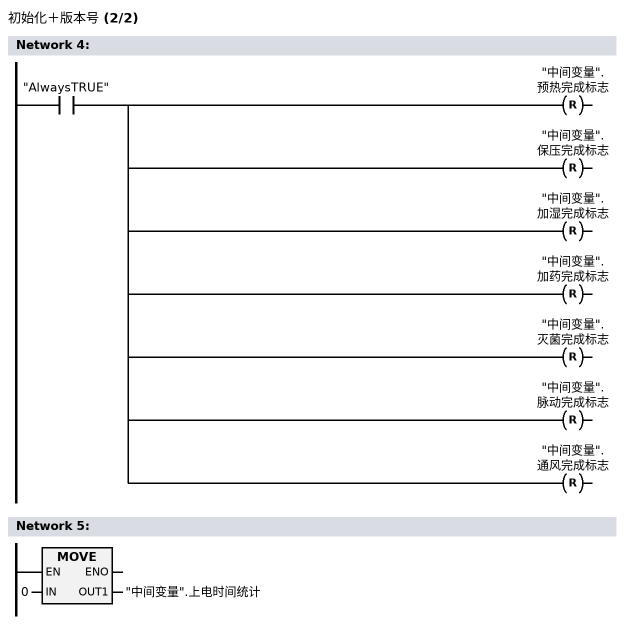
   RUNG wire#powerrail
      Contact( "AlwaysTRUE" )
      wire#w1
      R_Coil( "中间变量".预热完成标志 )
   END_RUNG
   RUNG wire#w1
      R_Coil( "中间变量".保压完成标志 )
   END_RUNG
   RUNG wire#w1
      R_Coil( "中间变量".加湿完成标志 )
   END_RUNG
   RUNG wire#w1
      R_Coil( "中间变量".加药完成标志 )
   END_RUNG
   RUNG wire#w1
      R_Coil( "中间变量".灭菌完成标志 )
   END_RUNG
   RUNG wire#w1
      R_Coil( "中间变量".脉动完成标志 )
   END_RUNG
   RUNG wire#w1
      R_Coil( "中间变量".通风完成标志 )
   END_RUNG
   // the same network as SCL:
   IF "AlwaysTRUE" THEN
       "中间变量".预热完成标志 := FALSE;
       "中间变量".保压完成标志 := FALSE;
       "中间变量".加湿完成标志 := FALSE;
       "中间变量".加药完成标志 := FALSE;
       "中间变量".灭菌完成标志 := FALSE;
       "中间变量".脉动完成标志 := FALSE;
       "中间变量".通风完成标志 := FALSE;
   END_IF;
END_REGION

REGION Network 5
   RUNG wire#powerrail
      Move(in := 0, out1 => "中间变量".上电时间统计)
   END_RUNG
   // the same network as SCL:
   "中间变量".上电时间统计 := 0;
END_REGION
END_FUNCTION

// folder: 101中间变量

FUNCTION_BLOCK "中间转换变量"   // FB4, LAD
{ S7_Optimized_Access := 'TRUE' }
VERSION : 0.1
   VAR RETAIN
      中间1 : Int;
      中间2 : Int;
      中间3 : Int;
      回空超时计算 : DInt;
      加药平衡时间计算 : DInt;
   END_VAR
BEGIN

REGION Network 1
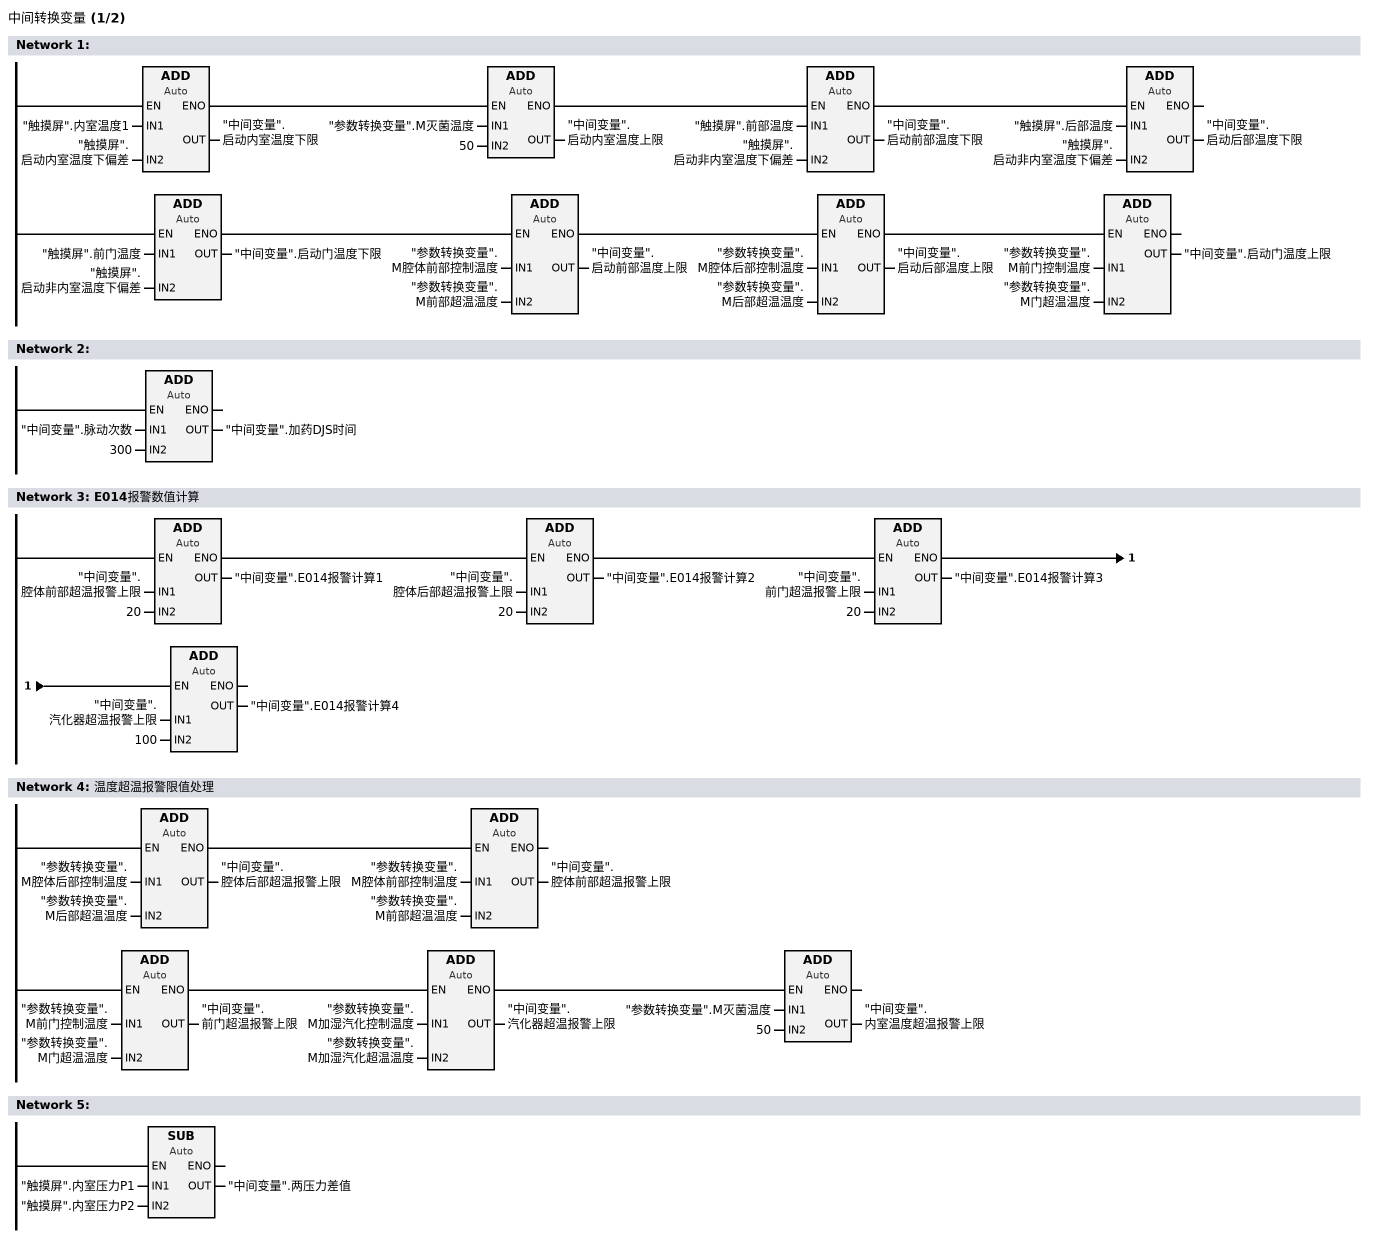
   RUNG wire#powerrail
      Add(in1 := "触摸屏".内室温度1, in2 := "触摸屏".启动内室温度下偏差, out => "中间变量".启动内室温度下限)
      Add(in1 := "参数转换变量".M灭菌温度, in2 := 50, out => "中间变量".启动内室温度上限)
      Add(in1 := "触摸屏".前部温度, in2 := "触摸屏".启动非内室温度下偏差, out => "中间变量".启动前部温度下限)
      Add(in1 := "触摸屏".后部温度, in2 := "触摸屏".启动非内室温度下偏差, out => "中间变量".启动后部温度下限)
   END_RUNG
   RUNG wire#powerrail
      Add(in1 := "触摸屏".前门温度, in2 := "触摸屏".启动非内室温度下偏差, out => "中间变量".启动门温度下限)
      Add(in1 := "参数转换变量".M腔体前部控制温度, in2 := "参数转换变量".M前部超温温度, out => "中间变量".启动前部温度上限)
      Add(in1 := "参数转换变量".M腔体后部控制温度, in2 := "参数转换变量".M后部超温温度, out => "中间变量".启动后部温度上限)
      Add(in1 := "参数转换变量".M前门控制温度, in2 := "参数转换变量".M门超温温度, out => "中间变量".启动门温度上限)
   END_RUNG
   // the same network as SCL:
   "中间变量".启动内室温度下限 := "触摸屏".内室温度1 + "触摸屏".启动内室温度下偏差;
   "中间变量".启动内室温度上限 := "参数转换变量".M灭菌温度 + 50;
   "中间变量".启动前部温度下限 := "触摸屏".前部温度 + "触摸屏".启动非内室温度下偏差;
   "中间变量".启动后部温度下限 := "触摸屏".后部温度 + "触摸屏".启动非内室温度下偏差;
   "中间变量".启动门温度下限 := "触摸屏".前门温度 + "触摸屏".启动非内室温度下偏差;
   "中间变量".启动前部温度上限 := "参数转换变量".M腔体前部控制温度 + "参数转换变量".M前部超温温度;
   "中间变量".启动后部温度上限 := "参数转换变量".M腔体后部控制温度 + "参数转换变量".M后部超温温度;
   "中间变量".启动门温度上限 := "参数转换变量".M前门控制温度 + "参数转换变量".M门超温温度;
END_REGION

REGION Network 2
   RUNG wire#powerrail
      Add(in1 := "中间变量".脉动次数, in2 := 300, out => "中间变量".加药DJS时间)
   END_RUNG
   // the same network as SCL:
   "中间变量".加药DJS时间 := "中间变量".脉动次数 + 300;
END_REGION

REGION Network 3: E014报警数值计算
   RUNG wire#powerrail
      Add(in1 := "中间变量".腔体前部超温报警上限, in2 := 20, out => "中间变量".E014报警计算1)
      Add(in1 := "中间变量".腔体后部超温报警上限, in2 := 20, out => "中间变量".E014报警计算2)
      Add(in1 := "中间变量".前门超温报警上限, in2 := 20, out => "中间变量".E014报警计算3)
      Add(in1 := "中间变量".汽化器超温报警上限, in2 := 100, out => "中间变量".E014报警计算4)
   END_RUNG
   // the same network as SCL:
   "中间变量".E014报警计算1 := "中间变量".腔体前部超温报警上限 + 20;
   "中间变量".E014报警计算2 := "中间变量".腔体后部超温报警上限 + 20;
   "中间变量".E014报警计算3 := "中间变量".前门超温报警上限 + 20;
   "中间变量".E014报警计算4 := "中间变量".汽化器超温报警上限 + 100;
END_REGION

REGION Network 4: 温度超温报警限值处理
   RUNG wire#powerrail
      Add(in1 := "参数转换变量".M腔体后部控制温度, in2 := "参数转换变量".M后部超温温度, out => "中间变量".腔体后部超温报警上限)
      Add(in1 := "参数转换变量".M腔体前部控制温度, in2 := "参数转换变量".M前部超温温度, out => "中间变量".腔体前部超温报警上限)
   END_RUNG
   RUNG wire#powerrail
      Add(in1 := "参数转换变量".M前门控制温度, in2 := "参数转换变量".M门超温温度, out => "中间变量".前门超温报警上限)
      Add(in1 := "参数转换变量".M加湿汽化控制温度, in2 := "参数转换变量".M加湿汽化超温温度, out => "中间变量".汽化器超温报警上限)
      Add(in1 := "参数转换变量".M灭菌温度, in2 := 50, out => "中间变量".内室温度超温报警上限)
   END_RUNG
   // the same network as SCL:
   "中间变量".腔体后部超温报警上限 := "参数转换变量".M腔体后部控制温度 + "参数转换变量".M后部超温温度;
   "中间变量".腔体前部超温报警上限 := "参数转换变量".M腔体前部控制温度 + "参数转换变量".M前部超温温度;
   "中间变量".前门超温报警上限 := "参数转换变量".M前门控制温度 + "参数转换变量".M门超温温度;
   "中间变量".汽化器超温报警上限 := "参数转换变量".M加湿汽化控制温度 + "参数转换变量".M加湿汽化超温温度;
   "中间变量".内室温度超温报警上限 := "参数转换变量".M灭菌温度 + 50;
END_REGION

REGION Network 5
   RUNG wire#powerrail
      Sub(in1 := "触摸屏".内室压力P1, in2 := "触摸屏".内室压力P2, out => "中间变量".两压力差值)
   END_RUNG
   // the same network as SCL:
   "中间变量".两压力差值 := "触摸屏".内室压力P1 - "触摸屏".内室压力P2;
END_REGION

REGION Network 6: 后门停止加热其中一个条件
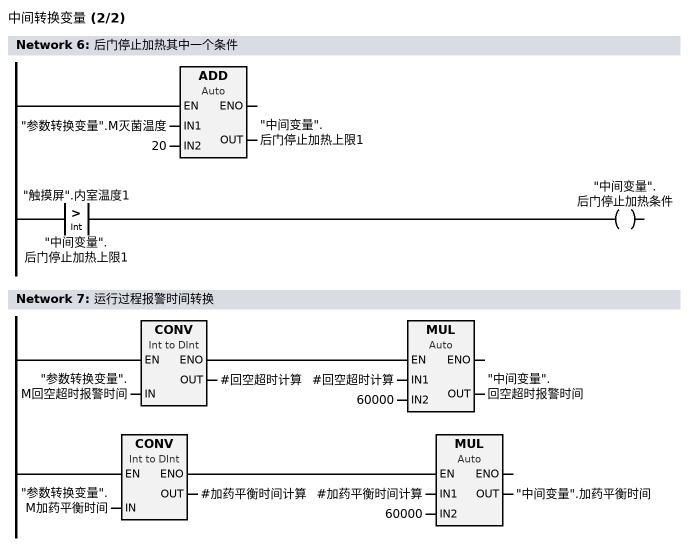
   RUNG wire#powerrail
      Add(in1 := "参数转换变量".M灭菌温度, in2 := 20, out => "中间变量".后门停止加热上限1)
   END_RUNG
   RUNG wire#powerrail
      { S7_Templates := "SrcType := Int" } GT_Contact(in1 := "触摸屏".内室温度1, in2 := "中间变量".后门停止加热上限1)
      Coil( "中间变量".后门停止加热条件 )
   END_RUNG
   // the same network as SCL:
   "中间变量".后门停止加热上限1 := "参数转换变量".M灭菌温度 + 20;
   "中间变量".后门停止加热条件 := "触摸屏".内室温度1 > "中间变量".后门停止加热上限1;
END_REGION

REGION Network 7: 运行过程报警时间转换
   RUNG wire#powerrail
      { S7_Templates := "[SrcType := Int, DestType := DInt]" } Convert(in := "参数转换变量".M回空超时报警时间, out => #回空超时计算)
      Mul(in1 := #回空超时计算, in2 := 60000, out => "中间变量".回空超时报警时间)
   END_RUNG
   RUNG wire#powerrail
      { S7_Templates := "[SrcType := Int, DestType := DInt]" } Convert(in := "参数转换变量".M加药平衡时间, out => #加药平衡时间计算)
      Mul(in1 := #加药平衡时间计算, in2 := 60000, out => "中间变量".加药平衡时间)
   END_RUNG
   // the same network as SCL:
   #回空超时计算 := INT_TO_DINT("参数转换变量".M回空超时报警时间);
   "中间变量".回空超时报警时间 := #回空超时计算 * 60000;
   #加药平衡时间计算 := INT_TO_DINT("参数转换变量".M加药平衡时间);
   "中间变量".加药平衡时间 := #加药平衡时间计算 * 60000;
END_REGION
END_FUNCTION_BLOCK

// folder: 12门功能控制

FUNCTION_BLOCK "门控制逻辑"   // FB14, LAD
{ S7_Optimized_Access := 'TRUE' }
VERSION : 0.1
   VAR_INPUT
      启动信号 : Bool;
      操作门开位 : Bool;
      操作门关位 : Bool;
      操作门障碍 : Bool;
      开操作门机械按钮 : Bool;
      关操作门机械按钮 : Bool;
      开操作门触摸按钮 : Bool;
      关操作门触摸按钮 : Bool;
      脚踢开关 : Bool;
      急停按钮 : Bool;
      内室压力符合标志 : Bool;
      程序运行标志 : Bool;
      门电机保护信号 : Bool;
      双门互锁功能开关 : Bool;
      对门关位 : Bool;
      操作门最大开启时间秒 : UInt;
      操作门最大关闭时间秒 : UInt;
      报警开关 : Word;
   END_VAR
   VAR_OUTPUT
      门状态 : UInt;
      报警码 : Word;
   END_VAR
   VAR
      机械开门按钮沿存储 : Bool;
      机械开门按钮状态 : Bool;
      触摸开门按钮沿存储 : Bool;
      触摸开门按钮状态 : Bool;
      机械关门按钮沿存储 : Bool;
      机械关门按钮状态 : Bool;
      触摸关门按钮沿存储 : Bool;
      触摸关门按钮状态 : Bool;
      脚踢开关沿存储 : Bool;
      脚踢开关状态 : Bool;
      开启操作门指令触发 : Bool;
      关闭操作门指令触发 : Bool;
      开门时间统计 : UInt;
      关门时间统计 : UInt;
      开门时间统计沿 : Bool;
      关门时间统计沿 : Bool;
      关闭门失败后需要开门标志 : Bool;
      门关闭失败重新开门等待时间 : UInt;
      门关闭失败重新开门时间统计沿 : Bool;
      报警码缓存 : Word;
      报警码输出时间统计 : UInt;
      报警码输出时间统计沿 : Bool;
      同时检测到门开位和关位信号时间统计 : UInt;
      同时检测到门开关位时间统计沿 : Bool;
      脚踢开关持续时间统计 : UInt;
      脚踢开关持续时间沿 : Bool;
   END_VAR
   VAR_TEMP
      操作门开启条件 : Bool;
      操作门关闭条件 : Bool;
      操作门最大开启时间 : UInt;
      操作门最大关闭时间 : UInt;
   END_VAR
   VAR_TEMP   // added for the SCL form of the ladder/FBD networks
      _w1 : Bool;
      _w2 : Bool;
      _w3 : Bool;
      _w4 : Bool;
      _w5 : Bool;
   END_VAR
BEGIN

REGION Network 1: 程序块初始化
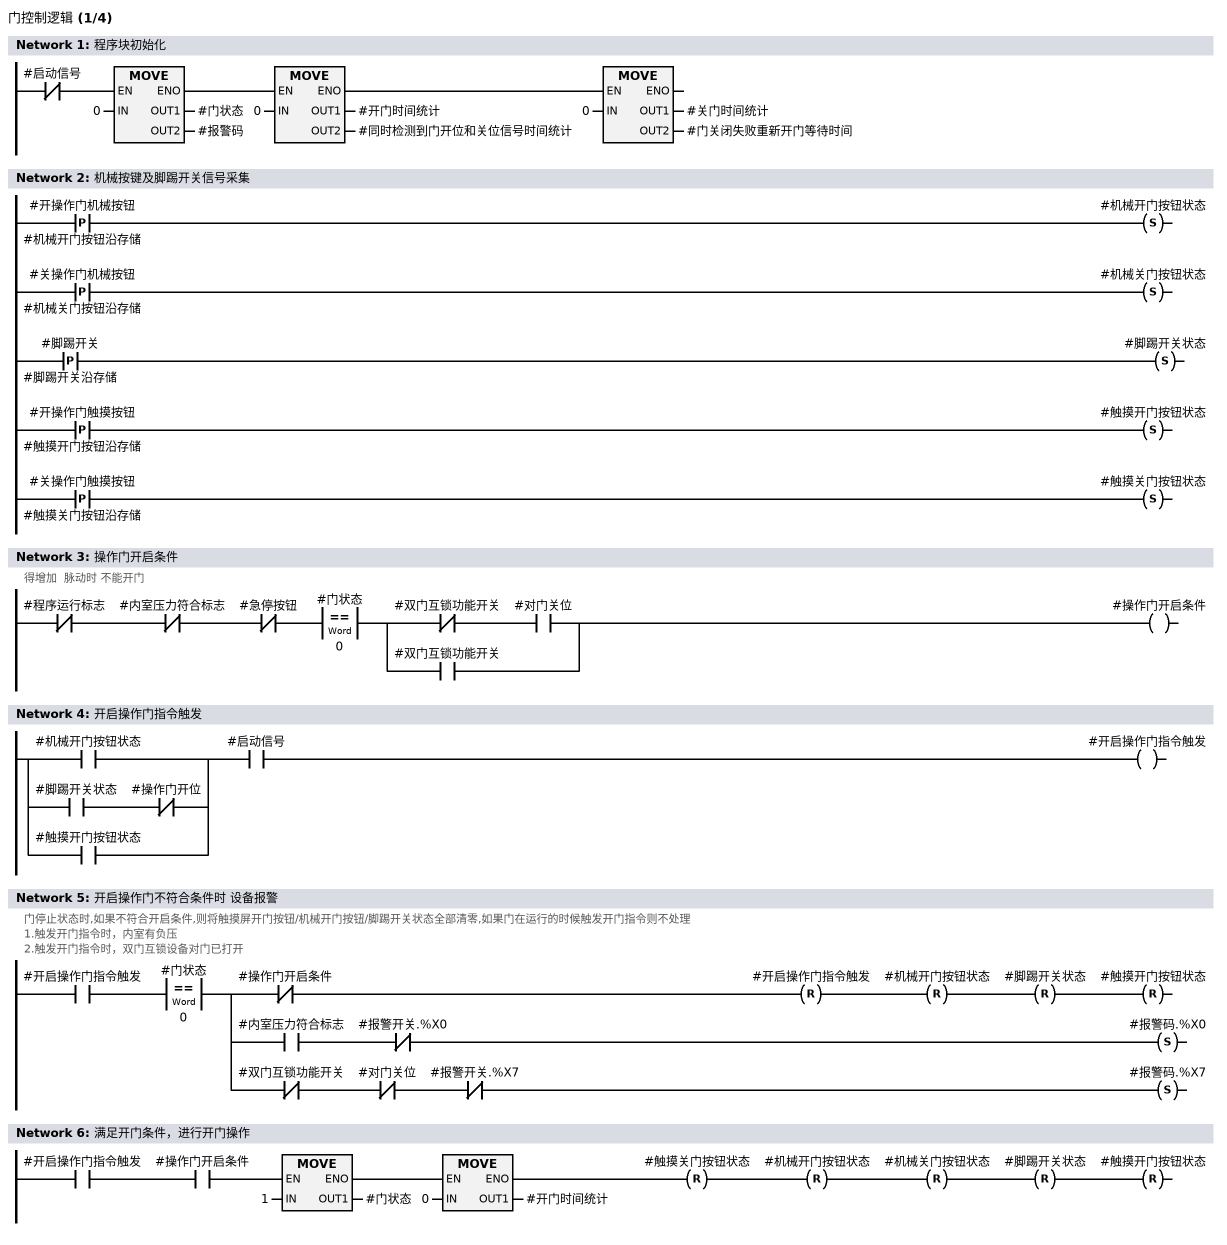
   RUNG wire#powerrail
      I_Contact( #启动信号 )
      Move(in := 0, out1 => #门状态, out2 => #报警码)
      Move(in := 0, out1 => #开门时间统计, out2 => #同时检测到门开位和关位信号时间统计)
      Move(in := 0, out1 => #关门时间统计, out2 => #门关闭失败重新开门等待时间)
   END_RUNG
   // the same network as SCL:
   IF NOT #启动信号 THEN
       #门状态 := 0;
       #报警码 := 0;
       #开门时间统计 := 0;
       #同时检测到门开位和关位信号时间统计 := 0;
       #关门时间统计 := 0;
       #门关闭失败重新开门等待时间 := 0;
   END_IF;
END_REGION

REGION Network 2: 机械按键及脚踢开关信号采集
   RUNG wire#powerrail
      P_Contact(operand := #开操作门机械按钮, bit := #机械开门按钮沿存储)
      S_Coil( #机械开门按钮状态 )
   END_RUNG
   RUNG wire#powerrail
      P_Contact(operand := #关操作门机械按钮, bit := #机械关门按钮沿存储)
      S_Coil( #机械关门按钮状态 )
   END_RUNG
   RUNG wire#powerrail
      P_Contact(operand := #脚踢开关, bit := #脚踢开关沿存储)
      S_Coil( #脚踢开关状态 )
   END_RUNG
   RUNG wire#powerrail
      P_Contact(operand := #开操作门触摸按钮, bit := #触摸开门按钮沿存储)
      S_Coil( #触摸开门按钮状态 )
   END_RUNG
   RUNG wire#powerrail
      P_Contact(operand := #关操作门触摸按钮, bit := #触摸关门按钮沿存储)
      S_Coil( #触摸关门按钮状态 )
   END_RUNG
   // the same network as SCL:
   #_w1 := #开操作门机械按钮 AND NOT #机械开门按钮沿存储;   // rising edge of #开操作门机械按钮
   #机械开门按钮沿存储 := #开操作门机械按钮;
   IF #_w1 THEN #机械开门按钮状态 := TRUE; END_IF;
   #_w2 := #关操作门机械按钮 AND NOT #机械关门按钮沿存储;   // rising edge of #关操作门机械按钮
   #机械关门按钮沿存储 := #关操作门机械按钮;
   IF #_w2 THEN #机械关门按钮状态 := TRUE; END_IF;
   #_w3 := #脚踢开关 AND NOT #脚踢开关沿存储;   // rising edge of #脚踢开关
   #脚踢开关沿存储 := #脚踢开关;
   IF #_w3 THEN #脚踢开关状态 := TRUE; END_IF;
   #_w4 := #开操作门触摸按钮 AND NOT #触摸开门按钮沿存储;   // rising edge of #开操作门触摸按钮
   #触摸开门按钮沿存储 := #开操作门触摸按钮;
   IF #_w4 THEN #触摸开门按钮状态 := TRUE; END_IF;
   #_w5 := #关操作门触摸按钮 AND NOT #触摸关门按钮沿存储;   // rising edge of #关操作门触摸按钮
   #触摸关门按钮沿存储 := #关操作门触摸按钮;
   IF #_w5 THEN #触摸关门按钮状态 := TRUE; END_IF;
END_REGION

REGION Network 3: 操作门开启条件
   // 得增加  脉动时 不能开门
   RUNG wire#powerrail
      I_Contact( #程序运行标志 )
      I_Contact( #内室压力符合标志 )
      I_Contact( #急停按钮 )
      { S7_Templates := "SrcType := Word" } EQ_Contact(in1 := #门状态, in2 := 0)
      wire#w1
      I_Contact( #双门互锁功能开关 )
      Contact( #对门关位 )
      wire#w2
      Coil( #操作门开启条件 )
   END_RUNG
   RUNG wire#w1
      Contact( #双门互锁功能开关 )
   END_RUNG wire#w2
   // the same network as SCL:
   #操作门开启条件 := NOT #程序运行标志 AND NOT #内室压力符合标志 AND NOT #急停按钮 AND (#门状态 = 0) AND ((NOT #双门互锁功能开关 AND #对门关位) OR #双门互锁功能开关);
END_REGION

REGION Network 4: 开启操作门指令触发
   RUNG wire#powerrail
      Contact( #机械开门按钮状态 )
      wire#w1
      Contact( #启动信号 )
      Coil( #开启操作门指令触发 )
   END_RUNG
   RUNG wire#powerrail
      Contact( #脚踢开关状态 )
      I_Contact( #操作门开位 )
   END_RUNG wire#w1
   RUNG wire#powerrail
      Contact( #触摸开门按钮状态 )
   END_RUNG wire#w1
   // the same network as SCL:
   #开启操作门指令触发 := (#机械开门按钮状态 OR (#脚踢开关状态 AND NOT #操作门开位) OR #触摸开门按钮状态) AND #启动信号;
END_REGION

REGION Network 5: 开启操作门不符合条件时 设备报警
   // 门停止状态时,如果不符合开启条件,则将触摸屏开门按钮/机械开门按钮/脚踢开关状态全部清零,如果门在运行的时候触发开门指令则不处理
   // 1.触发开门指令时，内室有负压  
   // 2.触发开门指令时，双门互锁设备对门已打开
   RUNG wire#powerrail
      Contact( #开启操作门指令触发 )
      { S7_Templates := "SrcType := Word" } EQ_Contact(in1 := #门状态, in2 := 0)
      wire#w1
      I_Contact( #操作门开启条件 )
      R_Coil( #开启操作门指令触发 )
      R_Coil( #机械开门按钮状态 )
      R_Coil( #脚踢开关状态 )
      R_Coil( #触摸开门按钮状态 )
   END_RUNG
   RUNG wire#w1
      Contact( #内室压力符合标志 )
      I_Contact( #报警开关.%X0 )
      S_Coil( #报警码.%X0 )
   END_RUNG
   RUNG wire#w1
      I_Contact( #双门互锁功能开关 )
      I_Contact( #对门关位 )
      I_Contact( #报警开关.%X7 )
      S_Coil( #报警码.%X7 )
   END_RUNG
   // the same network as SCL:
   #_w1 := #开启操作门指令触发 AND (#门状态 = 0);
   IF #_w1 AND NOT #操作门开启条件 THEN
       #开启操作门指令触发 := FALSE;
       #机械开门按钮状态 := FALSE;
       #脚踢开关状态 := FALSE;
       #触摸开门按钮状态 := FALSE;
   END_IF;
   IF #_w1 AND #内室压力符合标志 AND NOT #报警开关.%X0 THEN #报警码.%X0 := TRUE; END_IF;
   IF #_w1 AND NOT #双门互锁功能开关 AND NOT #对门关位 AND NOT #报警开关.%X7 THEN #报警码.%X7 := TRUE; END_IF;
END_REGION

REGION Network 6: 满足开门条件，进行开门操作
   RUNG wire#powerrail
      Contact( #开启操作门指令触发 )
      Contact( #操作门开启条件 )
      Move(in := 1, out1 => #门状态)
      Move(in := 0, out1 => #开门时间统计)
      R_Coil( #触摸关门按钮状态 )
      R_Coil( #机械开门按钮状态 )
      R_Coil( #机械关门按钮状态 )
      R_Coil( #脚踢开关状态 )
      R_Coil( #触摸开门按钮状态 )
   END_RUNG
   // the same network as SCL:
   IF #开启操作门指令触发 AND #操作门开启条件 THEN
       #门状态 := 1;
       #开门时间统计 := 0;
       #触摸关门按钮状态 := FALSE;
       #机械开门按钮状态 := FALSE;
       #机械关门按钮状态 := FALSE;
       #脚踢开关状态 := FALSE;
       #触摸开门按钮状态 := FALSE;
   END_IF;
END_REGION

REGION Network 7: 开操作门时间统计
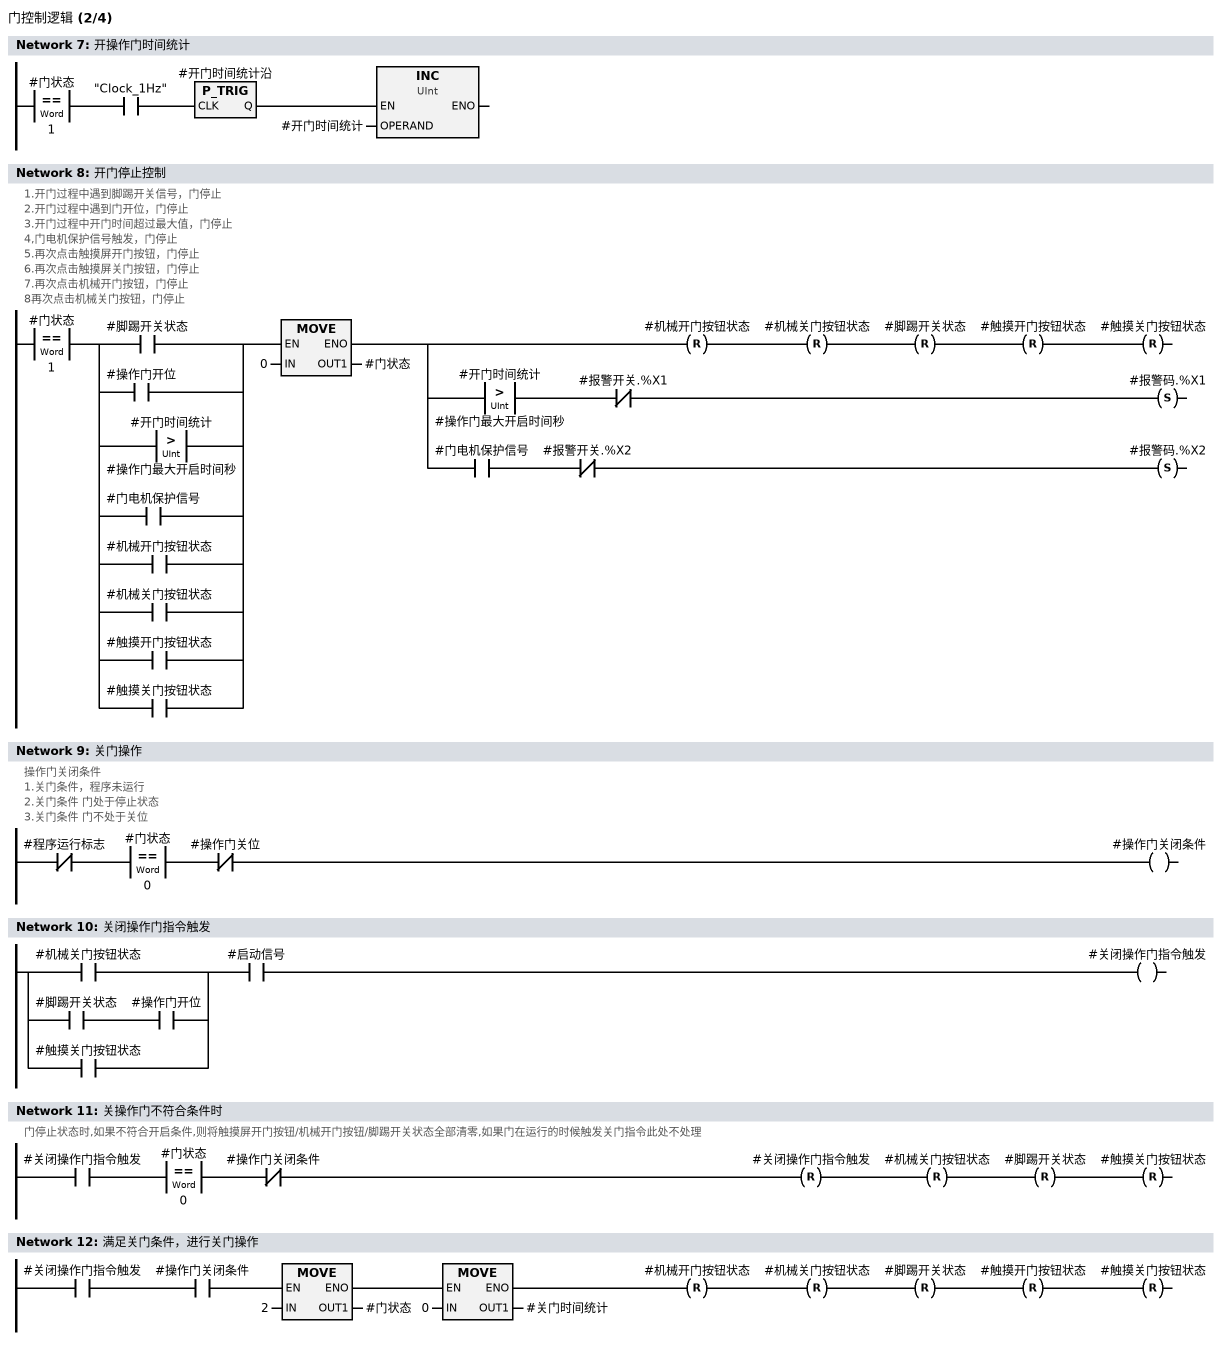
   RUNG wire#powerrail
      { S7_Templates := "SrcType := Word" } EQ_Contact(in1 := #门状态, in2 := 1)
      Contact( "Clock_1Hz" )
      P_Trig( #开门时间统计沿 )
      { S7_Templates := "DestType := UInt" } Inc( #开门时间统计 )
   END_RUNG
   // the same network as SCL:
   #_w1 := (#门状态 = 1) AND "Clock_1Hz";
   #_w2 := #_w1 AND NOT #开门时间统计沿;   // rising edge
   #开门时间统计沿 := #_w1;
   IF #_w2 THEN #开门时间统计 := #开门时间统计 + 1; END_IF;
END_REGION

REGION Network 8: 开门停止控制
   // 1.开门过程中遇到脚踢开关信号，门停止
   // 2.开门过程中遇到门开位，门停止
   // 3.开门过程中开门时间超过最大值，门停止
   // 4,门电机保护信号触发，门停止
   // 5.再次点击触摸屏开门按钮，门停止
   // 6.再次点击触摸屏关门按钮，门停止
   // 7.再次点击机械开门按钮，门停止
   // 8再次点击机械关门按钮，门停止
   RUNG wire#powerrail
      { S7_Templates := "SrcType := Word" } EQ_Contact(in1 := #门状态, in2 := 1)
      wire#w1
      Contact( #脚踢开关状态 )
      wire#w2
      Move(in := 0, out1 => #门状态)
      wire#w3
      R_Coil( #机械开门按钮状态 )
      R_Coil( #机械关门按钮状态 )
      R_Coil( #脚踢开关状态 )
      R_Coil( #触摸开门按钮状态 )
      R_Coil( #触摸关门按钮状态 )
   END_RUNG
   RUNG wire#w1
      Contact( #操作门开位 )
   END_RUNG wire#w2
   RUNG wire#w1
      { S7_Templates := "SrcType := UInt" } GT_Contact(in1 := #开门时间统计, in2 := #操作门最大开启时间秒)
   END_RUNG wire#w2
   RUNG wire#w1
      Contact( #门电机保护信号 )
   END_RUNG wire#w2
   RUNG wire#w1
      Contact( #机械开门按钮状态 )
   END_RUNG wire#w2
   RUNG wire#w1
      Contact( #机械关门按钮状态 )
   END_RUNG wire#w2
   RUNG wire#w1
      Contact( #触摸开门按钮状态 )
   END_RUNG wire#w2
   RUNG wire#w1
      Contact( #触摸关门按钮状态 )
   END_RUNG wire#w2
   RUNG wire#w3
      { S7_Templates := "SrcType := UInt" } GT_Contact(in1 := #开门时间统计, in2 := #操作门最大开启时间秒)
      I_Contact( #报警开关.%X1 )
      S_Coil( #报警码.%X1 )
   END_RUNG
   RUNG wire#w3
      Contact( #门电机保护信号 )
      I_Contact( #报警开关.%X2 )
      S_Coil( #报警码.%X2 )
   END_RUNG
   // the same network as SCL:
   #_w1 := (#门状态 = 1) AND (#脚踢开关状态 OR #操作门开位 OR (#开门时间统计 > #操作门最大开启时间秒) OR #门电机保护信号 OR #机械开门按钮状态 OR #机械关门按钮状态 OR #触摸开门按钮状态 OR #触摸关门按钮状态);
   IF #_w1 THEN
       #门状态 := 0;
       #机械开门按钮状态 := FALSE;
       #机械关门按钮状态 := FALSE;
       #脚踢开关状态 := FALSE;
       #触摸开门按钮状态 := FALSE;
       #触摸关门按钮状态 := FALSE;
   END_IF;
   IF #_w1 AND (#开门时间统计 > #操作门最大开启时间秒) AND NOT #报警开关.%X1 THEN #报警码.%X1 := TRUE; END_IF;
   IF #_w1 AND #门电机保护信号 AND NOT #报警开关.%X2 THEN #报警码.%X2 := TRUE; END_IF;
END_REGION

REGION Network 9: 关门操作
   // 操作门关闭条件
   // 1.关门条件，程序未运行
   // 2.关门条件 门处于停止状态
   // 3.关门条件 门不处于关位
   RUNG wire#powerrail
      I_Contact( #程序运行标志 )
      { S7_Templates := "SrcType := Word" } EQ_Contact(in1 := #门状态, in2 := 0)
      I_Contact( #操作门关位 )
      Coil( #操作门关闭条件 )
   END_RUNG
   // the same network as SCL:
   #操作门关闭条件 := NOT #程序运行标志 AND (#门状态 = 0) AND NOT #操作门关位;
END_REGION

REGION Network 10: 关闭操作门指令触发
   RUNG wire#powerrail
      Contact( #机械关门按钮状态 )
      wire#w1
      Contact( #启动信号 )
      Coil( #关闭操作门指令触发 )
   END_RUNG
   RUNG wire#powerrail
      Contact( #脚踢开关状态 )
      Contact( #操作门开位 )
   END_RUNG wire#w1
   RUNG wire#powerrail
      Contact( #触摸关门按钮状态 )
   END_RUNG wire#w1
   // the same network as SCL:
   #关闭操作门指令触发 := (#机械关门按钮状态 OR (#脚踢开关状态 AND #操作门开位) OR #触摸关门按钮状态) AND #启动信号;
END_REGION

REGION Network 11: 关操作门不符合条件时
   // 门停止状态时,如果不符合开启条件,则将触摸屏开门按钮/机械开门按钮/脚踢开关状态全部清零,如果门在运行的时候触发关门指令此处不处理
   RUNG wire#powerrail
      Contact( #关闭操作门指令触发 )
      { S7_Templates := "SrcType := Word" } EQ_Contact(in1 := #门状态, in2 := 0)
      I_Contact( #操作门关闭条件 )
      R_Coil( #关闭操作门指令触发 )
      R_Coil( #机械关门按钮状态 )
      R_Coil( #脚踢开关状态 )
      R_Coil( #触摸关门按钮状态 )
   END_RUNG
   // the same network as SCL:
   #_w1 := #关闭操作门指令触发 AND (#门状态 = 0) AND NOT #操作门关闭条件;
   IF #_w1 THEN
       #关闭操作门指令触发 := FALSE;
       #机械关门按钮状态 := FALSE;
       #脚踢开关状态 := FALSE;
       #触摸关门按钮状态 := FALSE;
   END_IF;
END_REGION

REGION Network 12: 满足关门条件，进行关门操作
   RUNG wire#powerrail
      Contact( #关闭操作门指令触发 )
      Contact( #操作门关闭条件 )
      Move(in := 2, out1 => #门状态)
      Move(in := 0, out1 => #关门时间统计)
      R_Coil( #机械开门按钮状态 )
      R_Coil( #机械关门按钮状态 )
      R_Coil( #脚踢开关状态 )
      R_Coil( #触摸开门按钮状态 )
      R_Coil( #触摸关门按钮状态 )
   END_RUNG
   // the same network as SCL:
   IF #关闭操作门指令触发 AND #操作门关闭条件 THEN
       #门状态 := 2;
       #关门时间统计 := 0;
       #机械开门按钮状态 := FALSE;
       #机械关门按钮状态 := FALSE;
       #脚踢开关状态 := FALSE;
       #触摸开门按钮状态 := FALSE;
       #触摸关门按钮状态 := FALSE;
   END_IF;
END_REGION

REGION Network 13: 关门动作时间统计
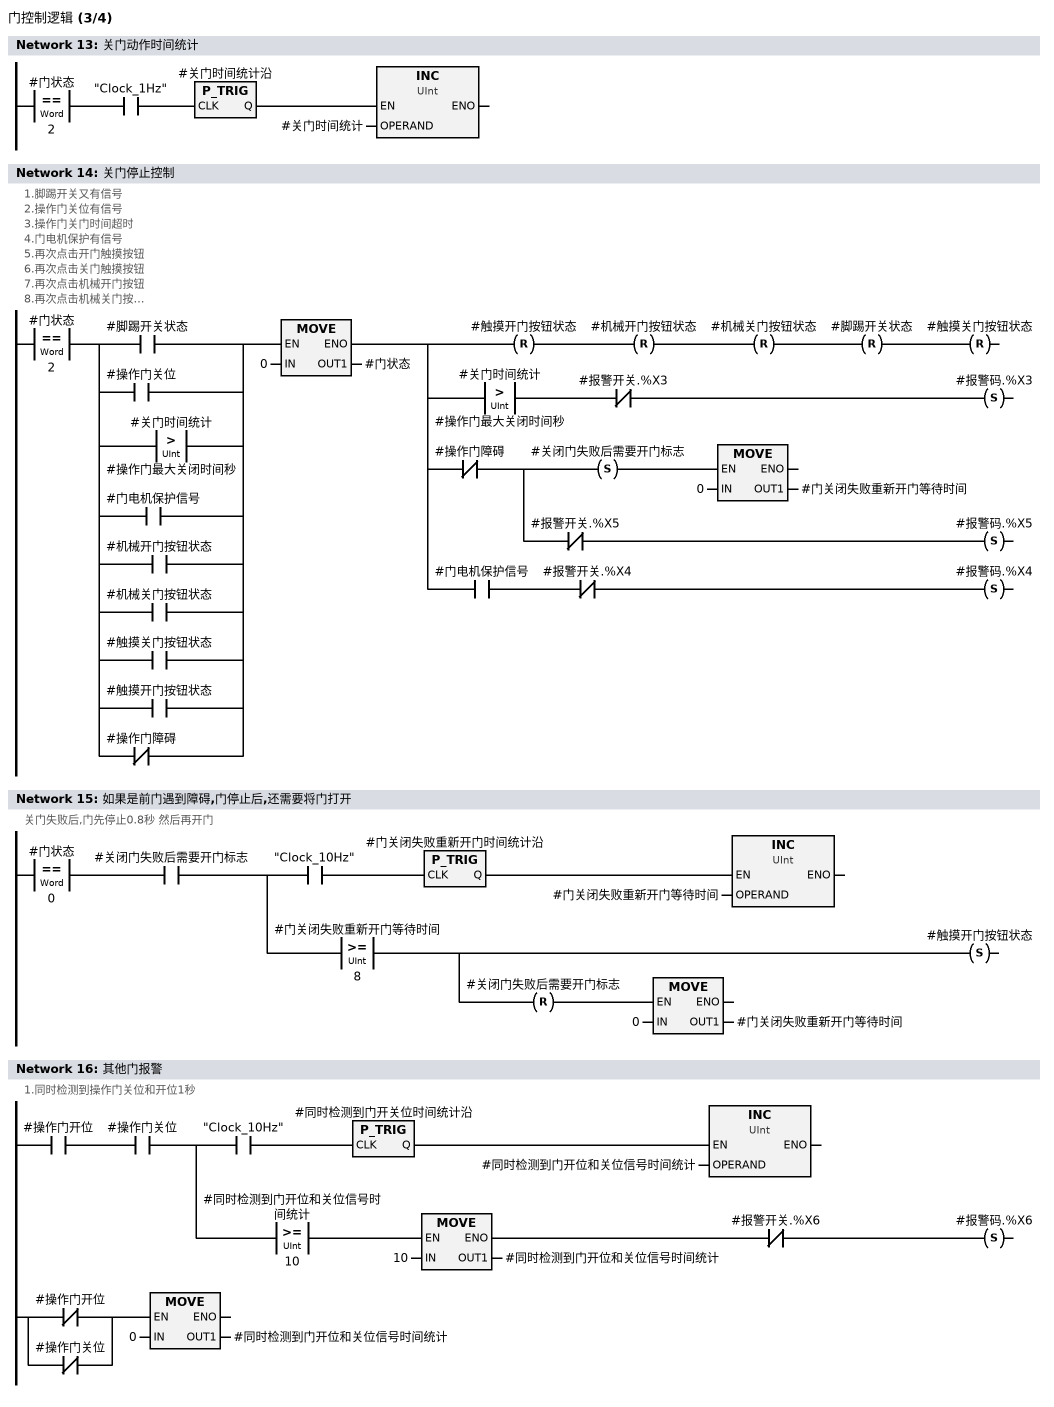
   RUNG wire#powerrail
      { S7_Templates := "SrcType := Word" } EQ_Contact(in1 := #门状态, in2 := 2)
      Contact( "Clock_1Hz" )
      P_Trig( #关门时间统计沿 )
      { S7_Templates := "DestType := UInt" } Inc( #关门时间统计 )
   END_RUNG
   // the same network as SCL:
   #_w1 := (#门状态 = 2) AND "Clock_1Hz";
   #_w2 := #_w1 AND NOT #关门时间统计沿;   // rising edge
   #关门时间统计沿 := #_w1;
   IF #_w2 THEN #关门时间统计 := #关门时间统计 + 1; END_IF;
END_REGION

